(* IEC 61131-3 sources: STEPROBOT/docs/plc_fixed_job_v1_2/现场升级_20261117, 10 files *)

(* ---- GVL_FileBridge.st ---- *)
{attribute 'qualified_only'}
VAR_GLOBAL PERSISTENT RETAIN
    (* Reserve these MW ranges in the FIELD project before importing. *)
    aCommand AT %MW6000 : ARRAY[0..119] OF WORD;
    aHeartbeat AT %MW6120 : ARRAY[0..4] OF WORD;
    aStatus AT %MW6200 : ARRAY[0..63] OF WORD;
END_VAR
VAR_GLOBAL
    (* LOCAL configuration only. Never map credentials/permit to Modbus. *)
    xFileTransferPermit : BOOL := FALSE;
    xReset : BOOL := FALSE;
    sFtpUser : STRING(64) := '';
    sFtpPassword : STRING(64) := '';
    aBuffer : ARRAY[0..1048575] OF BYTE;
    (* One-time LOCAL commissioning: exact existing project already bound to these three GDI numbers.
       This mode reuses bindings. It never edits robot system configuration. *)
    xFixedMappingConfirmed : BOOL := TRUE;
    sFixedProject : STRING(64) := 'pcjob_20261116_201104_7f547f98.sr';
    uiFixedCapture : UINT := UINT#1;
    uiFixedPath : UINT := UINT#2;
    uiFixedReturn : UINT := UINT#3;
    (* Nonretained: a reboot or failed update never authorizes a partly updated project. *)
    xFixedUpdateBusy : BOOL;
    xFixedReady : BOOL;
    xFixedIdle : BOOL;
END_VAR

(* ---- GVL_FileBridgeRetain.st ---- *)
{attribute 'qualified_only'}
VAR_GLOBAL PERSISTENT RETAIN
    udiBootCounter : UDINT := UDINT#0;
END_VAR

(* ---- GVL_RobotBridge.st ---- *)
{attribute 'qualified_only'}
VAR_GLOBAL PERSISTENT RETAIN
    // PC <-> PLC. Inovance native Modbus TCP slave: MWn <-> HR offset n.
    // Commission by reading HR300=16#4D42 and HR301=2 before permitting motion.
    aHostCmd AT %MW200 : ARRAY[0..15] OF WORD;
    aHostStatus AT %MW300 : ARRAY[0..63] OF WORD;

END_VAR

VAR_GLOBAL
    // PLC master -> STEP slave: FC04 / offset 0 / 32 WORD.
    aRobotRx : ARRAY[0..31] OF WORD;
    // PLC master -> STEP slave: ONE FC16 / offset 0 / 2 WORDs.
    // Map BOTH aRobotTx[0] and aRobotTx[1], NOT wRobotTxControl alone.
    aRobotTx : ARRAY[0..1] OF WORD;
    wRobotTxControl : WORD; // first-word diagnostic alias, not a separate channel

    // Local commissioning/operation inputs. Do not map these into aHostCmd.
    xCommissioned : BOOL := FALSE;
    // Set locally ONLY after checking DI49..56 and the GDI program bindings.
    xGdiProgramMappingConfirmed : BOOL := FALSE;
    xRemotePermit : BOOL := FALSE;
    // Optional native master/channel fault. FALSE leaves DO42 watchdog in use.
    xNativeModbusError : BOOL := FALSE;

    // Published live diagnostics.
    xRobotLinkOK : BOOL;
    xRobotRunning : BOOL;
    xRobotPaused : BOOL;
    xRobotStopped : BOOL;
    xRobotEnabled : BOOL;
    xRobotAlarm : BOOL;
    xRobotEmergency : BOOL;
    xRobotExternalAuto : BOOL;
    xHostRegistered : BOOL;
    xHostAlive : BOOL;
    xBusy : BOOL;
    xStopInterlock : BOOL;
    xLoadOperatorConfirmed : BOOL;
    uiFixedJobGuardVersion : UINT;
END_VAR

(* ---- GVL_RobotBridgeRetain.st ---- *)
{attribute 'qualified_only'}
VAR_GLOBAL PERSISTENT RETAIN
    // Incremented on application initialization, not on every scan.
    // Also require a fresh registration; a cold reset can reset RETAIN memory.
    udiBootCounter : UDINT := 0;
END_VAR

(* ---- F_FileCrc32.st ---- *)
FUNCTION F_FileCrc32 : UDINT
VAR_INPUT
    pData : POINTER TO BYTE;
    uiCount : UINT;
    udiSeed : UDINT;
END_VAR
VAR
    udiCrc : UDINT;
    uiI : UINT;
    uiBit : UINT;
END_VAR
(* Running reflected CRC-32. Caller supplies initial FFFFFFFF and final XOR. *)
udiCrc := udiSeed;
IF uiCount > UINT#0 THEN
    FOR uiI := UINT#0 TO uiCount - UINT#1 DO
        udiCrc := udiCrc XOR BYTE_TO_UDINT(pData[uiI]);
        FOR uiBit := UINT#0 TO UINT#7 DO
            IF (udiCrc AND UDINT#1) <> UDINT#0 THEN
                udiCrc := SHR(udiCrc, 1) XOR UDINT#16#EDB88320;
            ELSE
                udiCrc := SHR(udiCrc, 1);
            END_IF;
        END_FOR;
    END_FOR;
END_IF;
F_FileCrc32 := udiCrc;
END_FUNCTION

(* ---- F_FileNameValid.st ---- *)
FUNCTION F_FileNameValid : BOOL
VAR_INPUT
    sName : STRING(64);
    xProject : BOOL;
END_VAR
VAR
    pName : POINTER TO BYTE;
    uiI : UINT;
    uiBaseLength : UINT;
    xValid : BOOL;
    xChar : BOOL;
END_VAR
(* Flat lowercase ASCII names; no slash, CR/LF, spaces, or extra dots. *)
xValid := FALSE;
uiBaseLength := UINT#0;
IF xProject THEN
    IF (LEFT(sName, 6) = 'pcjob_') AND (RIGHT(sName, 3) = '.sr')
        AND (LEN(sName) >= 12) AND (LEN(sName) <= 48) THEN
        uiBaseLength := INT_TO_UINT(LEN(sName)) - UINT#3;
    END_IF;
ELSE
    IF (LEN(sName) >= 5) AND (LEN(sName) <= 48) THEN
        IF (RIGHT(sName, 4) = '.srp') OR (RIGHT(sName, 4) = '.srd')
            OR (RIGHT(sName, 4) = '.txt') THEN
            uiBaseLength := INT_TO_UINT(LEN(sName)) - UINT#4;
        END_IF;
    END_IF;
END_IF;
IF uiBaseLength > UINT#0 THEN
    xValid := TRUE;
    pName := ADR(sName);
    FOR uiI := UINT#0 TO uiBaseLength - UINT#1 DO
        xChar := ((pName[uiI] >= BYTE#97) AND (pName[uiI] <= BYTE#122))
            OR ((pName[uiI] >= BYTE#48) AND (pName[uiI] <= BYTE#57))
            OR (pName[uiI] = BYTE#95);
        IF NOT xChar THEN xValid := FALSE; END_IF;
    END_FOR;
END_IF;
F_FileNameValid := xValid;
END_FUNCTION

(* ---- F_FixedFileValid.st ---- *)
FUNCTION F_FixedFileValid : BOOL
VAR_INPUT
    sName : STRING(64);
END_VAR
F_FixedFileValid := (sName = '_project.srd')
    OR (sName = 'capture_home.srp') OR (sName = 'capture_home.srd')
    OR (sName = 'helix_25mms.srp') OR (sName = 'helix_25mms.srd')
    OR (sName = 'go_home.srp') OR (sName = 'go_home.srd');
END_FUNCTION

(* ---- FB_FileFtp.st ---- *)
FUNCTION_BLOCK FB_FileFtp
VAR_INPUT
    xStart : BOOL;
    xAbort : BOOL;
    pBuffer : POINTER TO BYTE;
    udiSize : UDINT;
    sProject : STRING(64);
    sFile : STRING(64);
    xCreateProject : BOOL;
    xReplaceFixed : BOOL;
    sUser : STRING(64);
    sPassword : STRING(64);
END_VAR
VAR CONSTANT
    cdiControlID : DINT := DINT#245;
    cdiDataID : DINT := DINT#246;
END_VAR
VAR_OUTPUT
    xDone : BOOL := FALSE;
    xTestPassed : BOOL := FALSE;
    xError : BOOL := FALSE;
    xLoginOk : BOOL := FALSE;
    xBaseDirOk : BOOL := FALSE;
    xScratchCreated : BOOL := FALSE;
    xUploadComplete : BOOL := FALSE;
    xReadbackComplete : BOOL := FALSE;
    xContentMatch : BOOL := FALSE;
    xQuitOk : BOOL := FALSE;
    xCleanupOk : BOOL := FALSE;
    uiStep : UINT := UINT#0;
    uiErrorStage : UINT := UINT#0;
    wErrorID : WORD := WORD#0;
    wDataCloseErrorID : WORD := WORD#0;
    wControlCloseErrorID : WORD := WORD#0;
    udiExpectedBytes : UDINT := UDINT#0;
    udiUploadedBytes : UDINT := UDINT#0;
    udiReadbackBytes : UDINT := UDINT#0;
    uiReplyCode : UINT := UINT#0;
    uiUserReplyCode : UINT := UINT#0;
    uiPassReplyCode : UINT := UINT#0;
    uiBaseDirReplyCode : UINT := UINT#0;
    uiNameCheckReplyCode : UINT := UINT#0;
    uiMkdReplyCode : UINT := UINT#0;
    uiStorReplyCode : UINT := UINT#0;
    uiUploadCompleteCode : UINT := UINT#0;
    uiRetrReplyCode : UINT := UINT#0;
    uiDownloadCompleteCode : UINT := UINT#0;
    uiPasvPort : UINT := UINT#0;
    wReadbackEndStatus : WORD := WORD#0;
    sRemotePath : STRING(160);
    sLastReply : STRING(255);
    sMkdReply : STRING(255);
    sPasvReply : STRING(255);
    sUploadReply : STRING(255);
    sDownloadReply : STRING(255);
    xControlOwned : BOOL := FALSE;
    xDataOwned : BOOL := FALSE;
    xUploadDataConnected : BOOL := FALSE;
    xDownloadDataConnected : BOOL := FALSE;
    xLineTruncated : BOOL := FALSE;

END_VAR
VAR
    (* Caller owns immutable buffer until xDone and clean socket closure. *)
    xAbortLatched : BOOL;
    xProgress : BOOL;
    xDirectoryReady : BOOL;
    xReplaceRun : BOOL;
    sFileRun : STRING(64);
    pBufferRun : POINTER TO BYTE;

    stControlServer : CmpHCTCPIP.ADDRESS := (strIPAddr := '192.168.3.188', uiPort := UINT#21);
    stDataServer : CmpHCTCPIP.ADDRESS;
    fbControlClient : CmpHCTCPIP.SktTCPClient;
    fbControlReceive : CmpHCTCPIP.SktTCPRecv;
    fbControlSend : CmpHCTCPIP.SktTCPSend;
    fbControlClose : CmpHCTCPIP.SktClose;
    fbDataClient : CmpHCTCPIP.SktTCPClient;
    fbDataSend : CmpHCTCPIP.SktTCPSend;
    fbDataReceive : CmpHCTCPIP.SktTCPRecv;
    fbDataClose : CmpHCTCPIP.SktClose;
    fbReplyTimeout : TON;
    fbCommandTimeout : TON;
    fbUploadTimeout : TON;
    fbReadbackTimeout : TON;
    fbDataCloseTimeout : TON;
    fbControlCloseTimeout : TON;

    xStartOld : BOOL := FALSE;
    xFail : BOOL := FALSE;
    xFinishedNow : BOOL := FALSE;
    wPendingError : WORD := WORD#0;
    uiPendingStage : UINT := UINT#0;
    uiPhase : UINT := UINT#0;
    uiNextCommand : UINT := UINT#0;
    uiTransferMode : UINT := UINT#0;
    xReplyReady : BOOL := FALSE;
    xReplyAccepted : BOOL := FALSE;
    xDigits : BOOL := FALSE;
    xMultiline : BOOL := FALSE;
    sMultilineCode : STRING(3);
    sLine : STRING(255);
    pLine : POINTER TO BYTE;
    uiLineLength : UINT := UINT#0;
    aControlRx : ARRAY[0..0] OF BYTE;
    sCommand : STRING(160);
    pCommand : POINTER TO BYTE;
    uiCommandIndex : UINT := UINT#0;
    uiCommandLength : UINT := UINT#0;
    aControlTx : ARRAY[0..0] OF BYTE;
    aDataTx : ARRAY[0..0] OF BYTE;
    aDataRx : ARRAY[0..0] OF BYTE;
    sUserRun : STRING(64);
    sPasswordRun : STRING(64);
    sScratchRun : STRING(64);
    pCredential : POINTER TO BYTE;
    uiI : UINT := UINT#0;
    xNameCharacter : BOOL := FALSE;
    xBytesMatch : BOOL := FALSE;
    xReadbackEndCandidate : BOOL := FALSE;
    xDataCloseFailed : BOOL := FALSE;
    pReply : POINTER TO BYTE;
    aPasv : ARRAY[0..5] OF UINT;
    uiPasvField : UINT := UINT#0;
    uiPasvValue : UINT := UINT#0;
    xPasvValid : BOOL := FALSE;
    xPasvInTuple : BOOL := FALSE;
    xPasvClosed : BOOL := FALSE;
    xPasvHasDigit : BOOL := FALSE;
END_VAR
(* Derived from field-passed PRG_FtpUploadProbe. New bridge is NOT field validated. *)
(* IDs 245/246 must be free; default cabinet 192.168.3.188:21. *)
(* One-byte send/reset preserves the tested Socket behavior. No motion commands. *)
pLine := ADR(sLine);
pCommand := ADR(sCommand);
xFail := FALSE;
xFinishedNow := FALSE;
xReplyReady := FALSE;
wPendingError := WORD#0;
uiPendingStage := UINT#20 + uiPhase * UINT#10;

IF uiStep = UINT#40 THEN
    aControlTx[0] := pCommand[uiCommandIndex];
END_IF;
IF uiStep = UINT#60 THEN
    IF udiUploadedBytes < udiExpectedBytes THEN
        aDataTx[0] := pBufferRun[udiUploadedBytes];
    END_IF;
END_IF;

fbControlClient(xExecute := uiStep = UINT#10, diConnectID := cdiControlID,
    stServerAddress := stControlServer);
fbControlReceive(xEnable := uiStep = UINT#20, diConnectID := cdiControlID,
    abyData := aControlRx, uiDataSize := UINT#1);
fbControlSend(xExecute := uiStep = UINT#40, diConnectID := cdiControlID,
    abyData := aControlTx, uiDataSize := UINT#1, uiTimeOut := UINT#1000);
fbDataClient(xExecute := uiStep = UINT#50, diConnectID := cdiDataID,
    stServerAddress := stDataServer);
fbDataSend(xExecute := uiStep = UINT#60, diConnectID := cdiDataID,
    abyData := aDataTx, uiDataSize := UINT#1, uiTimeOut := UINT#1000);
fbDataReceive(xEnable := uiStep = UINT#70, diConnectID := cdiDataID,
    abyData := aDataRx, uiDataSize := UINT#1);
fbDataClose(xExecute := ((uiStep = UINT#80) OR (uiStep = UINT#90))
    AND xDataOwned AND NOT xDataCloseFailed, diConnectID := cdiDataID);
fbControlClose(xExecute := (uiStep = UINT#95) AND xControlOwned,
    diConnectID := cdiControlID);
fbReplyTimeout(IN := uiStep = UINT#20, PT := T#20s);
fbCommandTimeout(IN := (uiStep = UINT#40) OR (uiStep = UINT#45), PT := T#30s);
xProgress := ((uiStep = UINT#60) AND fbDataSend.xDone)
    OR ((uiStep = UINT#70) AND (fbDataReceive.uiCount > UINT#0));
fbUploadTimeout(IN := ((uiStep = UINT#60) OR (uiStep = UINT#65)) AND NOT xProgress,
    PT := T#30s);
fbReadbackTimeout(IN := (uiStep = UINT#70) AND NOT xProgress, PT := T#30s);
fbDataCloseTimeout(IN := ((uiStep = UINT#80) OR (uiStep = UINT#90))
    AND xDataOwned AND NOT xDataCloseFailed, PT := T#5s);
fbControlCloseTimeout(IN := uiStep = UINT#95, PT := T#5s);

(* Bounded control-reply parser; identical-code SPACE terminates multiline replies. *)
IF (uiStep = UINT#20) AND NOT fbControlReceive.xError THEN
    IF fbControlReceive.uiCount > UINT#0 THEN
        IF aControlRx[0] = BYTE#10 THEN
            IF uiLineLength > UINT#0 THEN
                IF pLine[uiLineLength - UINT#1] = BYTE#13 THEN
                    uiLineLength := uiLineLength - UINT#1;
                    pLine[uiLineLength] := BYTE#0;
                END_IF;
            END_IF;
            IF xMultiline THEN
                IF LEFT(sLine, 4) = CONCAT(sMultilineCode, ' ') THEN
                    xMultiline := FALSE;
                    xReplyReady := TRUE;
                END_IF;
            ELSE
                xDigits := FALSE;
                IF uiLineLength >= UINT#4 THEN
                    xDigits := (pLine[0] >= BYTE#48) AND (pLine[0] <= BYTE#57)
                        AND (pLine[1] >= BYTE#48) AND (pLine[1] <= BYTE#57)
                        AND (pLine[2] >= BYTE#48) AND (pLine[2] <= BYTE#57);
                END_IF;
                IF xDigits THEN
                    IF pLine[3] = BYTE#45 THEN
                        xMultiline := TRUE;
                        sMultilineCode := LEFT(sLine, 3);
                    ELSIF pLine[3] = BYTE#32 THEN
                        xReplyReady := TRUE;
                    ELSE
                        xFail := TRUE;
                        wPendingError := WORD#16#F203;
                    END_IF;
                ELSE
                    xFail := TRUE;
                    wPendingError := WORD#16#F203;
                END_IF;
            END_IF;
            IF xReplyReady THEN
                uiReplyCode := (BYTE_TO_UINT(pLine[0]) - UINT#48) * UINT#100
                    + (BYTE_TO_UINT(pLine[1]) - UINT#48) * UINT#10
                    + BYTE_TO_UINT(pLine[2]) - UINT#48;
                sLastReply := sLine;
            ELSIF xFail THEN
                sLastReply := sLine;
            END_IF;
            sLine := '';
            uiLineLength := UINT#0;
        ELSE
            IF uiLineLength < UINT#255 THEN
                pLine[uiLineLength] := aControlRx[0];
                uiLineLength := uiLineLength + UINT#1;
                pLine[uiLineLength] := BYTE#0;
            ELSE
                xLineTruncated := TRUE;
                sLastReply := sLine;
                xFail := TRUE;
                wPendingError := WORD#16#F204;
            END_IF;
        END_IF;
    END_IF;
END_IF;

CASE uiStep OF
    UINT#0:
        IF xStart AND NOT xStartOld THEN
            xAbortLatched := FALSE;
            xDirectoryReady := FALSE;
            xDone := FALSE;
            xTestPassed := FALSE;
            xError := FALSE;
            xLoginOk := FALSE;
            xBaseDirOk := FALSE;
            xScratchCreated := FALSE;
            xUploadComplete := FALSE;
            xReadbackComplete := FALSE;
            xContentMatch := FALSE;
            xQuitOk := FALSE;
            xCleanupOk := FALSE;
            xUploadDataConnected := FALSE;
            xDownloadDataConnected := FALSE;
            xDataCloseFailed := FALSE;
            xLineTruncated := FALSE;
            xReadbackEndCandidate := FALSE;
            xBytesMatch := TRUE;
            uiErrorStage := UINT#0;
            wErrorID := WORD#0;
            wDataCloseErrorID := WORD#0;
            wControlCloseErrorID := WORD#0;
            wReadbackEndStatus := WORD#0;
            udiUploadedBytes := UDINT#0;
            udiReadbackBytes := UDINT#0;
            uiReplyCode := UINT#0;
            uiUserReplyCode := UINT#0;
            uiPassReplyCode := UINT#0;
            uiBaseDirReplyCode := UINT#0;
            uiNameCheckReplyCode := UINT#0;
            uiMkdReplyCode := UINT#0;
            uiStorReplyCode := UINT#0;
            uiUploadCompleteCode := UINT#0;
            uiRetrReplyCode := UINT#0;
            uiDownloadCompleteCode := UINT#0;
            uiPasvPort := UINT#0;
            sLastReply := '';
            sMkdReply := '';
            sPasvReply := '';
            sUploadReply := '';
            sDownloadReply := '';
            sLine := '';
            uiLineLength := UINT#0;
            xMultiline := FALSE;
            sMultilineCode := '';
            uiPhase := UINT#0;
            uiTransferMode := UINT#0;
            sUserRun := sUser;
            sPasswordRun := sPassword;
            sScratchRun := sProject;
            sFileRun := sFile;
            xReplaceRun := xReplaceFixed;
            pBufferRun := pBuffer;
            sRemotePath := CONCAT(CONCAT(CONCAT('/UserPrograms/', sScratchRun), '/'), sFileRun);
            udiExpectedBytes := udiSize;
            uiPendingStage := UINT#1;
            IF (LEN(sUserRun) = 0) OR (LEN(sPasswordRun) = 0) THEN
                xFail := TRUE;
                wPendingError := WORD#16#F200;
            ELSE
                pCredential := ADR(sUserRun);
                FOR uiI := UINT#0 TO INT_TO_UINT(LEN(sUserRun)) - UINT#1 DO
                    IF (pCredential[uiI] < BYTE#32) OR (pCredential[uiI] > BYTE#126) THEN
                        xFail := TRUE;
                        wPendingError := WORD#16#F207;
                    END_IF;
                END_FOR;
                pCredential := ADR(sPasswordRun);
                FOR uiI := UINT#0 TO INT_TO_UINT(LEN(sPasswordRun)) - UINT#1 DO
                    IF (pCredential[uiI] < BYTE#32) OR (pCredential[uiI] > BYTE#126) THEN
                        xFail := TRUE;
                        wPendingError := WORD#16#F207;
                    END_IF;
                END_FOR;
            END_IF;
            IF NOT F_FileNameValid(sScratchRun, TRUE)
                OR NOT F_FileNameValid(sFileRun, FALSE)
                OR (udiExpectedBytes > UDINT#1048576)
                OR (pBufferRun = 0) THEN
                xFail := TRUE;
                wPendingError := WORD#16#F209;
            END_IF;
            IF xReplaceRun AND (NOT GVL_FileBridge.xFixedMappingConfirmed
                OR (GVL_RobotBridge.uiFixedJobGuardVersion <> UINT#120)
                OR NOT GVL_FileBridge.xFixedIdle OR (sScratchRun <> GVL_FileBridge.sFixedProject)
                OR NOT F_FixedFileValid(sFileRun)) THEN
                xFail := TRUE;
                wPendingError := WORD#16#F20C;
            END_IF;
            IF NOT xFail THEN
                uiStep := UINT#10;
            END_IF;
        END_IF;

    UINT#10:
        IF fbControlClient.xError THEN
            xFail := TRUE;
            wPendingError := fbControlClient.wErrorID;
            uiPendingStage := UINT#10;
        ELSIF fbControlClient.xDone THEN
            xControlOwned := TRUE;
            uiStep := UINT#20;
        END_IF;

    UINT#20:
        IF fbControlReceive.xError THEN
            xFail := TRUE;
            wPendingError := fbControlReceive.wErrorID;
        ELSIF NOT xFail THEN
            IF xReplyReady THEN
                xReplyAccepted := FALSE;
                CASE uiPhase OF
                    UINT#0:
                        IF uiReplyCode = UINT#220 THEN
                            xReplyAccepted := TRUE;
                            uiNextCommand := UINT#1;
                            uiStep := UINT#30;
                        ELSIF uiReplyCode = UINT#120 THEN
                            xReplyAccepted := TRUE;
                        END_IF;
                    UINT#1:
                        uiUserReplyCode := uiReplyCode;
                        IF uiReplyCode = UINT#331 THEN
                            xReplyAccepted := TRUE;
                            uiNextCommand := UINT#2;
                            uiStep := UINT#30;
                        ELSIF uiReplyCode = UINT#230 THEN
                            xReplyAccepted := TRUE;
                            xLoginOk := TRUE;
                            uiNextCommand := UINT#3;
                            uiStep := UINT#30;
                        END_IF;
                    UINT#2:
                        uiPassReplyCode := uiReplyCode;
                        IF uiReplyCode = UINT#230 THEN
                            xReplyAccepted := TRUE;
                            xLoginOk := TRUE;
                            uiNextCommand := UINT#3;
                            uiStep := UINT#30;
                        END_IF;
                    UINT#3:
                        uiBaseDirReplyCode := uiReplyCode;
                        IF uiReplyCode = UINT#250 THEN
                            xReplyAccepted := TRUE;
                            xBaseDirOk := TRUE;
                            IF xCreateProject OR xReplaceRun THEN
                                uiNextCommand := UINT#14;
                            ELSE
                                uiNextCommand := UINT#5;
                            END_IF;
                            uiStep := UINT#30;
                        END_IF;
                    UINT#14:
                        uiNameCheckReplyCode := uiReplyCode;
                        IF uiReplyCode = UINT#550 THEN
                            xReplyAccepted := TRUE;
                            IF xReplaceRun THEN
                                (* Fixed binding must already exist: never silently create another target. *)
                                xFail := TRUE;
                                wPendingError := WORD#16#F20B;
                            ELSE
                                uiNextCommand := UINT#4;
                                uiStep := UINT#30;
                            END_IF;
                        ELSIF uiReplyCode = UINT#250 THEN
                            xReplyAccepted := TRUE;
                            IF xReplaceRun THEN
                                xDirectoryReady := TRUE;
                                uiNextCommand := UINT#6;
                                uiStep := UINT#30;
                            ELSE
                                (* Original mode retains its no-overwrite behavior. *)
                                xFail := TRUE;
                                wPendingError := WORD#16#F208;
                            END_IF;
                        END_IF;
                    UINT#4:
                        uiMkdReplyCode := uiReplyCode;
                        sMkdReply := sLastReply;
                        IF uiReplyCode = UINT#257 THEN
                            xReplyAccepted := TRUE;
                            xScratchCreated := TRUE;
                            uiNextCommand := UINT#5;
                            uiStep := UINT#30;
                        END_IF;
                    UINT#5:
                        IF uiReplyCode = UINT#250 THEN
                            xDirectoryReady := TRUE;
                            xReplyAccepted := TRUE;
                            uiNextCommand := UINT#6;
                            uiStep := UINT#30;
                        END_IF;
                    UINT#6:
                        IF uiReplyCode = UINT#200 THEN
                            xReplyAccepted := TRUE;
                            uiNextCommand := UINT#7;
                            uiStep := UINT#30;
                        END_IF;
                    UINT#7, UINT#10:
                        IF uiReplyCode = UINT#227 THEN
                            xReplyAccepted := TRUE;
                            sPasvReply := sLastReply;
                            uiStep := UINT#35;
                        END_IF;
                    UINT#8:
                        uiStorReplyCode := uiReplyCode;
                        IF (uiReplyCode = UINT#125) OR (uiReplyCode = UINT#150) THEN
                            xReplyAccepted := TRUE;
                            IF udiExpectedBytes = UDINT#0 THEN
                                (* Empty STOR still needs data EOF, 226 and exact RETR. *)
                                uiStep := UINT#80;
                            ELSE
                                uiStep := UINT#60;
                            END_IF;
                        END_IF;
                    UINT#9:
                        uiUploadCompleteCode := uiReplyCode;
                        sUploadReply := sLastReply;
                        IF (uiReplyCode = UINT#226) OR (uiReplyCode = UINT#250) THEN
                            xReplyAccepted := TRUE;
                            xUploadComplete := TRUE;
                            uiNextCommand := UINT#10;
                            uiStep := UINT#30;
                        END_IF;
                    UINT#11:
                        uiRetrReplyCode := uiReplyCode;
                        IF (uiReplyCode = UINT#125) OR (uiReplyCode = UINT#150) THEN
                            xReplyAccepted := TRUE;
                            uiStep := UINT#70;
                        END_IF;
                    UINT#12:
                        uiDownloadCompleteCode := uiReplyCode;
                        sDownloadReply := sLastReply;
                        IF (uiReplyCode = UINT#226) OR (uiReplyCode = UINT#250) THEN
                            xReplyAccepted := TRUE;
                            xReadbackComplete := TRUE;
                            xContentMatch := xBytesMatch AND xReadbackEndCandidate
                                AND (udiReadbackBytes = udiExpectedBytes);
                            IF xContentMatch THEN
                                uiNextCommand := UINT#13;
                                uiStep := UINT#30;
                            ELSE
                                xFail := TRUE;
                                wPendingError := WORD#16#F205;
                            END_IF;
                        END_IF;
                    UINT#13:
                        IF uiReplyCode = UINT#221 THEN
                            xReplyAccepted := TRUE;
                            xQuitOk := TRUE;
                            uiStep := UINT#90;
                        END_IF;
                END_CASE;
                IF NOT xReplyAccepted THEN
                    xFail := TRUE;
                    wPendingError := WORD#16#F202;
                END_IF;
            ELSIF fbReplyTimeout.Q THEN
                xFail := TRUE;
                wPendingError := WORD#16#F201;
            END_IF;
        END_IF;

    UINT#30:
        uiPhase := uiNextCommand;
        CASE uiNextCommand OF
            UINT#1: sCommand := CONCAT(CONCAT('USER ', sUserRun), '$R$N');
            UINT#2: sCommand := CONCAT(CONCAT('PASS ', sPasswordRun), '$R$N');
            UINT#3: sCommand := 'CWD /UserPrograms$R$N';
            UINT#4: sCommand := CONCAT(CONCAT('MKD ', sScratchRun), '$R$N');
            UINT#5, UINT#14: sCommand := CONCAT(CONCAT('CWD ', sScratchRun), '$R$N');
            UINT#6: sCommand := 'TYPE I$R$N';
            UINT#7, UINT#10: sCommand := 'PASV$R$N';
            UINT#8: sCommand := CONCAT(CONCAT('STOR ', sFileRun), '$R$N');
            UINT#11: sCommand := CONCAT(CONCAT('RETR ', sFileRun), '$R$N');
            UINT#13: sCommand := 'QUIT$R$N';
        ELSE
            xFail := TRUE;
            wPendingError := WORD#16#F20A;
        END_CASE;
        IF NOT xFail THEN
            uiCommandLength := INT_TO_UINT(LEN(sCommand));
            uiCommandIndex := UINT#0;
            uiStep := UINT#40;
        END_IF;

    UINT#35:
        (* Parse six decimal octets in the first parenthesized PASV tuple. *)
        pReply := ADR(sPasvReply);
        xPasvValid := TRUE;
        xPasvInTuple := FALSE;
        xPasvClosed := FALSE;
        xPasvHasDigit := FALSE;
        uiPasvField := UINT#0;
        uiPasvValue := UINT#0;
        FOR uiI := UINT#0 TO INT_TO_UINT(LEN(sPasvReply)) - UINT#1 DO
            IF NOT xPasvInTuple THEN
                IF pReply[uiI] = BYTE#40 THEN
                    xPasvInTuple := TRUE;
                END_IF;
            ELSIF NOT xPasvClosed THEN
                IF (pReply[uiI] >= BYTE#48) AND (pReply[uiI] <= BYTE#57) THEN
                    xPasvHasDigit := TRUE;
                    IF uiPasvValue <= UINT#255 THEN
                        uiPasvValue := uiPasvValue * UINT#10 + BYTE_TO_UINT(pReply[uiI]) - UINT#48;
                        IF uiPasvValue > UINT#255 THEN
                            xPasvValid := FALSE;
                        END_IF;
                    ELSE
                        xPasvValid := FALSE;
                    END_IF;
                ELSIF (pReply[uiI] = BYTE#44) OR (pReply[uiI] = BYTE#41) THEN
                    IF NOT xPasvHasDigit OR (uiPasvField > UINT#5) OR (uiPasvValue > UINT#255) THEN
                        xPasvValid := FALSE;
                    ELSE
                        aPasv[uiPasvField] := uiPasvValue;
                        uiPasvField := uiPasvField + UINT#1;
                    END_IF;
                    uiPasvValue := UINT#0;
                    xPasvHasDigit := FALSE;
                    IF pReply[uiI] = BYTE#41 THEN
                        xPasvClosed := TRUE;
                    END_IF;
                ELSE
                    xPasvValid := FALSE;
                END_IF;
            END_IF;
        END_FOR;
        IF NOT xPasvInTuple OR NOT xPasvClosed OR (uiPasvField <> UINT#6) THEN
            xPasvValid := FALSE;
        END_IF;
        IF xPasvValid THEN
            uiPasvPort := aPasv[4] * UINT#256 + aPasv[5];
            IF (uiPasvPort = UINT#0) OR (uiPasvPort = UINT#21) THEN
                xPasvValid := FALSE;
            END_IF;
        END_IF;
        IF xPasvValid THEN
            (* Data connections are pinned to the control server, not a third-party PASV IP. *)
            stDataServer.strIPAddr := stControlServer.strIPAddr;
            stDataServer.uiPort := uiPasvPort;
            xDataCloseFailed := FALSE;
            IF uiPhase = UINT#7 THEN
                uiTransferMode := UINT#1;
            ELSE
                uiTransferMode := UINT#2;
            END_IF;
            uiStep := UINT#50;
        ELSE
            xFail := TRUE;
            wPendingError := WORD#16#F20B;
        END_IF;

    UINT#40:
        IF fbControlSend.xError THEN
            xFail := TRUE;
            wPendingError := fbControlSend.wErrorID;
        ELSIF fbControlSend.xDone THEN
            uiCommandIndex := uiCommandIndex + UINT#1;
            uiStep := UINT#45;
        ELSIF fbCommandTimeout.Q THEN
            xFail := TRUE;
            wPendingError := WORD#16#F206;
        END_IF;

    UINT#45:
        IF uiCommandIndex >= uiCommandLength THEN
            sCommand := '';
            aControlTx[0] := BYTE#0;
            sLine := '';
            uiLineLength := UINT#0;
            xMultiline := FALSE;
            sMultilineCode := '';
            uiStep := UINT#20;
        ELSIF fbCommandTimeout.Q THEN
            xFail := TRUE;
            wPendingError := WORD#16#F206;
        ELSE
            uiStep := UINT#40;
        END_IF;

    UINT#50:
        uiPendingStage := UINT#200 + uiTransferMode;
        IF fbDataClient.xError THEN
            xFail := TRUE;
            wPendingError := fbDataClient.wErrorID;
        ELSIF fbDataClient.xDone THEN
            xDataOwned := TRUE;
            IF uiTransferMode = UINT#1 THEN
                xUploadDataConnected := TRUE;
                uiNextCommand := UINT#8;
            ELSE
                xDownloadDataConnected := TRUE;
                uiNextCommand := UINT#11;
            END_IF;
            uiStep := UINT#30;
        END_IF;

    UINT#60:
        uiPendingStage := UINT#210;
        IF fbDataSend.xError THEN
            xFail := TRUE;
            wPendingError := fbDataSend.wErrorID;
        ELSIF fbDataSend.xDone THEN
            udiUploadedBytes := udiUploadedBytes + UDINT#1;
            uiStep := UINT#65;
        ELSIF fbUploadTimeout.Q THEN
            xFail := TRUE;
            wPendingError := WORD#16#F206;
        END_IF;

    UINT#65:
        uiPendingStage := UINT#210;
        IF udiUploadedBytes >= udiExpectedBytes THEN
            aDataTx[0] := BYTE#0;
            uiStep := UINT#80;
        ELSIF fbUploadTimeout.Q THEN
            xFail := TRUE;
            wPendingError := WORD#16#F206;
        ELSE
            uiStep := UINT#60;
        END_IF;

    UINT#70:
        uiPendingStage := UINT#220;
        IF fbDataReceive.xError THEN
            wReadbackEndStatus := fbDataReceive.wErrorID;
            (* In the supplied source, zero-length recv and recv failure share 0011. *)
            (* This is only an end candidate: exact bytes AND FTP completion are required. *)
            IF (wReadbackEndStatus = WORD#16#0011) AND xBytesMatch
                AND (udiReadbackBytes = udiExpectedBytes) THEN
                xReadbackEndCandidate := TRUE;
                uiStep := UINT#80;
            ELSE
                xFail := TRUE;
                wPendingError := fbDataReceive.wErrorID;
            END_IF;
        ELSIF fbDataReceive.uiCount > UINT#0 THEN
            IF udiReadbackBytes >= udiExpectedBytes THEN
                xBytesMatch := FALSE;
                xFail := TRUE;
                wPendingError := WORD#16#F205;
            ELSE
                IF aDataRx[0] <> pBufferRun[udiReadbackBytes] THEN
                    xBytesMatch := FALSE;
                    xFail := TRUE;
                    wPendingError := WORD#16#F205;
                END_IF;
                udiReadbackBytes := udiReadbackBytes + UDINT#1;
            END_IF;
        ELSIF fbReadbackTimeout.Q THEN
            xFail := TRUE;
            wPendingError := WORD#16#F201;
        END_IF;

    UINT#80:
        IF fbDataClose.xError OR fbDataCloseTimeout.Q THEN
            IF fbDataClose.xError THEN
                wDataCloseErrorID := fbDataClose.wErrorID;
            ELSE
                wDataCloseErrorID := WORD#16#F20C;
            END_IF;
            xDataCloseFailed := TRUE;
            IF NOT xError THEN
                xError := TRUE;
                wErrorID := wDataCloseErrorID;
                uiErrorStage := UINT#290;
            END_IF;
            uiStep := UINT#95;
        ELSIF fbDataClose.xDone THEN
            xDataOwned := FALSE;
            IF uiTransferMode = UINT#1 THEN
                uiPhase := UINT#9;
            ELSE
                uiPhase := UINT#12;
            END_IF;
            uiStep := UINT#20;
        END_IF;

    UINT#90:
        IF NOT xDataOwned OR xDataCloseFailed THEN
            uiStep := UINT#95;
        ELSIF fbDataClose.xError OR fbDataCloseTimeout.Q THEN
            IF fbDataClose.xError THEN
                wDataCloseErrorID := fbDataClose.wErrorID;
            ELSE
                wDataCloseErrorID := WORD#16#F20C;
            END_IF;
            xDataCloseFailed := TRUE;
            IF NOT xError THEN
                xError := TRUE;
                wErrorID := wDataCloseErrorID;
                uiErrorStage := UINT#290;
            END_IF;
            uiStep := UINT#95;
        ELSIF fbDataClose.xDone THEN
            xDataOwned := FALSE;
            uiStep := UINT#95;
        END_IF;

    UINT#95:
        IF NOT xControlOwned THEN
            xDone := TRUE;
            xFinishedNow := TRUE;
            uiStep := UINT#100;
        ELSIF fbControlClose.xError OR fbControlCloseTimeout.Q THEN
            IF fbControlClose.xError THEN
                wControlCloseErrorID := fbControlClose.wErrorID;
            ELSE
                wControlCloseErrorID := WORD#16#F20C;
            END_IF;
            IF NOT xError THEN
                xError := TRUE;
                wErrorID := wControlCloseErrorID;
                uiErrorStage := UINT#295;
            END_IF;
            xDone := TRUE;
            xFinishedNow := TRUE;
            uiStep := UINT#100;
        ELSIF fbControlClose.xDone THEN
            xControlOwned := FALSE;
            xDone := TRUE;
            xFinishedNow := TRUE;
            uiStep := UINT#100;
        END_IF;

    UINT#100:
        IF NOT xStart AND NOT xControlOwned AND NOT xDataOwned THEN
            uiStep := UINT#0;
        END_IF;
END_CASE;

(* Never cancel a pending native connect before its terminal result. *)
IF xAbort AND (uiStep <> UINT#0) AND (uiStep <> UINT#100) THEN
    xAbortLatched := TRUE;
END_IF;
IF xAbortLatched AND (uiStep <> UINT#0) AND (uiStep <> UINT#10)
    AND (uiStep <> UINT#50) AND (uiStep <> UINT#90)
    AND (uiStep <> UINT#95) AND (uiStep <> UINT#100) THEN
    xFail := TRUE;
    wPendingError := WORD#16#F20D;
END_IF;
IF xFail THEN
    IF NOT xError THEN
        xError := TRUE;
        wErrorID := wPendingError;
        uiErrorStage := uiPendingStage;
    END_IF;
    uiStep := UINT#90;
END_IF;

IF xFinishedNow THEN
    xCleanupOk := NOT xControlOwned AND NOT xDataOwned
        AND (wDataCloseErrorID = WORD#0) AND (wControlCloseErrorID = WORD#0);
    xTestPassed := xLoginOk AND xBaseDirOk AND xDirectoryReady
        AND xUploadDataConnected AND xDownloadDataConnected
        AND xUploadComplete AND xReadbackComplete AND xContentMatch
        AND xQuitOk AND xCleanupOk AND NOT xError;
    sPasswordRun := '';
    sUserRun := '';
    sCommand := '';
    aControlTx[0] := BYTE#0;
    aDataTx[0] := BYTE#0;
END_IF;
xStartOld := xStart;
END_FUNCTION_BLOCK

(* ---- PRG_FileBridge.st ---- *)
PROGRAM PRG_FileBridge
VAR
    xInit : BOOL;
    xResetOld : BOOL;
    aPrevious : ARRAY[0..119] OF WORD;
    aSeen : ARRAY[0..119] OF WORD;
    aFrame : ARRAY[0..119] OF WORD;
    aAccepted : ARRAY[0..119] OF WORD;
    aFrameBytes : ARRAY[0..235] OF BYTE;
    aPayload : ARRAY[0..191] OF BYTE;
    aNames : ARRAY[0..31] OF STRING(64);
    uiState : UINT;
    wError : WORD;
    udiOwner : UDINT;
    udiAck : UDINT;
    uiAckOp : UINT;
    udiSize : UDINT;
    udiReceived : UDINT;
    udiExpectedCrc : UDINT;
    udiRunningCrc : UDINT := UDINT#16#FFFFFFFF;
    udiTotalSize : UDINT;
    uiVerified : UINT;
    uiExpectedFiles : UINT;
    uiOrdinal : UINT;
    uiMode : UINT;
    sProject : STRING(64);
    sFile : STRING(64);
    fbFtp : FB_FileFtp;
    fbLease : TON;
    wHeartbeatOld : WORD;
    xKick : BOOL;
    xStable : BOOL;
    xNew : BOOL;
    xSame : BOOL;
    xAccept : BOOL;
    xActive : BOOL;
    xClean : BOOL;
    xFileVerified : BOOL;
    xFtpStarted : BOOL;
    wReject : WORD;
    udiRejectSeq : UDINT;
    udiRejectOwner : UDINT;
    wRequestError : WORD;
    udiSeq : UDINT;
    udiSession : UDINT;
    udiBoot : UDINT;
    udiFrameCrc : UDINT;
    udiFrameSize : UDINT;
    udiOffset : UDINT;
    udiFileCrc : UDINT;
    uiOp : UINT;
    uiLength : UINT;
    uiCount : UINT;
    uiIndex : UINT;
    uiField : UINT;
    uiPos : UINT;
    uiI : UINT;
    uiJ : UINT;
    uiSnapshot : UINT;
    wFlags : WORD;
    sNewProject : STRING(64);
    sNewFile : STRING(64);
    pName : POINTER TO BYTE;
    xNamesOk : BOOL;
    xPairsOk : BOOL;
    xFound : BOOL;
    xGlobal : BOOL;
    uiPrograms : UINT;
    sPair : STRING(64);
    sReadyProject : STRING(64);
    uiReadyCapture : UINT;
    uiReadyPath : UINT;
    uiReadyReturn : UINT;
    xFixedConfig : BOOL;
    udiFixedProjectCrc : UDINT;
    uiSessionCapture : UINT;
    uiSessionPath : UINT;
    uiSessionReturn : UINT;
END_VAR

(* This program NEVER writes robot motion/control outputs or GDI selection. *)
IF NOT xInit THEN
    GVL_FileBridge.xFixedReady := FALSE;
    GVL_FileBridge.xFixedUpdateBusy := FALSE;
    IF GVL_FileBridgeRetain.udiBootCounter = UDINT#16#FFFFFFFF THEN
        GVL_FileBridgeRetain.udiBootCounter := UDINT#1;
    ELSE
        GVL_FileBridgeRetain.udiBootCounter := GVL_FileBridgeRetain.udiBootCounter + UDINT#1;
    END_IF;
    FOR uiI := UINT#0 TO UINT#119 DO
        aPrevious[uiI] := GVL_FileBridge.aCommand[uiI];
        aSeen[uiI] := GVL_FileBridge.aCommand[uiI];
    END_FOR;
    xInit := TRUE;
END_IF;

xFixedConfig := GVL_FileBridge.xFixedMappingConfirmed
    AND (GVL_RobotBridge.uiFixedJobGuardVersion = UINT#120)
    AND F_FileNameValid(GVL_FileBridge.sFixedProject, TRUE)
    AND (GVL_FileBridge.uiFixedCapture >= UINT#1) AND (GVL_FileBridge.uiFixedCapture <= UINT#255)
    AND (GVL_FileBridge.uiFixedPath >= UINT#1) AND (GVL_FileBridge.uiFixedPath <= UINT#255)
    AND (GVL_FileBridge.uiFixedReturn >= UINT#1) AND (GVL_FileBridge.uiFixedReturn <= UINT#255)
    AND (GVL_FileBridge.uiFixedCapture <> GVL_FileBridge.uiFixedPath)
    AND (GVL_FileBridge.uiFixedCapture <> GVL_FileBridge.uiFixedReturn)
    AND (GVL_FileBridge.uiFixedPath <> GVL_FileBridge.uiFixedReturn);
GVL_FileBridge.xFixedIdle := GVL_RobotBridge.xRobotLinkOK AND GVL_RobotBridge.xRobotStopped
    AND NOT GVL_RobotBridge.xRobotRunning AND NOT GVL_RobotBridge.xRobotPaused
    AND NOT GVL_RobotBridge.xRobotEnabled AND NOT GVL_RobotBridge.xBusy;
IF NOT xFixedConfig OR (sReadyProject <> GVL_FileBridge.sFixedProject)
    OR (uiReadyCapture <> GVL_FileBridge.uiFixedCapture) OR (uiReadyPath <> GVL_FileBridge.uiFixedPath)
    OR (uiReadyReturn <> GVL_FileBridge.uiFixedReturn) THEN
    GVL_FileBridge.xFixedReady := FALSE;
END_IF;
udiFixedProjectCrc := F_FileCrc32(ADR(GVL_FileBridge.sFixedProject),
    INT_TO_UINT(LEN(GVL_FileBridge.sFixedProject)), UDINT#16#FFFFFFFF) XOR UDINT#16#FFFFFFFF;

xClean := NOT fbFtp.xControlOwned AND NOT fbFtp.xDataOwned
    AND ((fbFtp.uiStep = UINT#0) OR (fbFtp.uiStep = UINT#100));
IF GVL_FileBridge.xReset AND NOT xResetOld AND xClean
    AND (uiState <> UINT#300) AND (uiState <> UINT#310) THEN
    uiState := UINT#0;
    wError := WORD#0;
    udiOwner := UDINT#0;
    udiAck := UDINT#0;
    uiAckOp := UINT#0;
    uiVerified := UINT#0;
    uiExpectedFiles := UINT#0;
    udiReceived := UDINT#0;
    udiSize := UDINT#0;
    xFileVerified := FALSE;
    GVL_FileBridge.xFixedReady := FALSE;
    wReject := WORD#0;
END_IF;
xResetOld := GVL_FileBridge.xReset;

xActive := (uiState = UINT#100) OR (uiState = UINT#200)
    OR (uiState = UINT#300) OR (uiState = UINT#310);
xKick := FALSE;
IF (GVL_FileBridge.aHeartbeat[0] = UDINT_TO_WORD(SHR(udiOwner, 16)))
    AND (GVL_FileBridge.aHeartbeat[1] = UDINT_TO_WORD(udiOwner))
    AND (GVL_FileBridge.aHeartbeat[2] = UDINT_TO_WORD(SHR(GVL_FileBridgeRetain.udiBootCounter, 16)))
    AND (GVL_FileBridge.aHeartbeat[3] = UDINT_TO_WORD(GVL_FileBridgeRetain.udiBootCounter))
    AND (GVL_FileBridge.aHeartbeat[4] <> wHeartbeatOld) THEN
    wHeartbeatOld := GVL_FileBridge.aHeartbeat[4];
    xKick := TRUE;
END_IF;
fbLease(IN := xActive AND NOT xKick, PT := T#10s);

(* Two consecutive identical samples, then CRC of big-endian WORD bytes. *)
xStable := TRUE;
xNew := FALSE;
FOR uiI := UINT#0 TO UINT#119 DO
    aFrame[uiI] := GVL_FileBridge.aCommand[uiI];
    IF aFrame[uiI] <> aPrevious[uiI] THEN xStable := FALSE; END_IF;
    IF aFrame[uiI] <> aSeen[uiI] THEN xNew := TRUE; END_IF;
    aPrevious[uiI] := aFrame[uiI];
END_FOR;
IF xStable AND xNew THEN
    FOR uiI := UINT#0 TO UINT#119 DO aSeen[uiI] := aFrame[uiI]; END_FOR;
    FOR uiI := UINT#0 TO UINT#117 DO
        aFrameBytes[uiI * UINT#2] := WORD_TO_BYTE(SHR(aFrame[uiI], 8));
        aFrameBytes[uiI * UINT#2 + UINT#1] := WORD_TO_BYTE(aFrame[uiI] AND WORD#255);
    END_FOR;
    FOR uiI := UINT#0 TO UINT#95 DO
        aPayload[uiI * UINT#2] := WORD_TO_BYTE(SHR(aFrame[uiI + UINT#20], 8));
        aPayload[uiI * UINT#2 + UINT#1] := WORD_TO_BYTE(aFrame[uiI + UINT#20] AND WORD#255);
    END_FOR;
    uiOp := WORD_TO_UINT(aFrame[2]);
    udiSeq := SHL(WORD_TO_UDINT(aFrame[3]), 16) OR WORD_TO_UDINT(aFrame[4]);
    udiSession := SHL(WORD_TO_UDINT(aFrame[5]), 16) OR WORD_TO_UDINT(aFrame[6]);
    udiBoot := SHL(WORD_TO_UDINT(aFrame[7]), 16) OR WORD_TO_UDINT(aFrame[8]);
    udiFrameSize := SHL(WORD_TO_UDINT(aFrame[9]), 16) OR WORD_TO_UDINT(aFrame[10]);
    udiOffset := SHL(WORD_TO_UDINT(aFrame[11]), 16) OR WORD_TO_UDINT(aFrame[12]);
    uiLength := WORD_TO_UINT(aFrame[13]);
    udiFileCrc := SHL(WORD_TO_UDINT(aFrame[14]), 16) OR WORD_TO_UDINT(aFrame[15]);
    udiFrameCrc := F_FileCrc32(ADR(aFrameBytes), UINT#236, UDINT#16#FFFFFFFF) XOR UDINT#16#FFFFFFFF;
    wRequestError := WORD#0;
    xAccept := FALSE;
    IF (aFrame[0] <> WORD#16#F7B1) OR (aFrame[1] <> WORD#1)
        OR (aFrame[19] <> WORD#0) OR (aFrame[116] <> WORD#0) OR (aFrame[117] <> WORD#0)
        OR (uiLength > UINT#192) OR (udiSeq = UDINT#0) OR (udiSession = UDINT#0) THEN
        wRequestError := WORD#16#E001;
    ELSIF udiFrameCrc <> (SHL(WORD_TO_UDINT(aFrame[118]), 16) OR WORD_TO_UDINT(aFrame[119])) THEN
        wRequestError := WORD#16#E002;
    ELSIF udiBoot <> GVL_FileBridgeRetain.udiBootCounter THEN
        wRequestError := WORD#16#E003;
    ELSIF (udiSession = udiOwner) AND (udiSeq = udiAck) THEN
        xSame := TRUE;
        FOR uiI := UINT#0 TO UINT#119 DO
            IF aAccepted[uiI] <> aFrame[uiI] THEN xSame := FALSE; END_IF;
        END_FOR;
        IF NOT xSame THEN wRequestError := WORD#16#E004; END_IF;
        (* Exact replay: existing ACK/status only; NEVER repeat file/FTP operations. *)
    ELSE
        IF (uiOp = UINT#1) AND ((uiState = UINT#0) OR (uiState = UINT#400)) THEN
            IF (udiSeq <> UDINT#1) OR NOT xClean THEN wRequestError := WORD#16#E005; END_IF;
        ELSIF udiSession <> udiOwner THEN
            wRequestError := WORD#16#E006;
        ELSIF (udiSeq <= udiAck) OR (udiAck = UDINT#16#FFFFFFFF) THEN
            wRequestError := WORD#16#E005;
        ELSIF (uiOp <> UINT#4) AND (uiOp <> UINT#6) AND (udiSeq <> udiAck + UDINT#1) THEN
            wRequestError := WORD#16#E005;
        END_IF;
        IF NOT GVL_FileBridge.xFileTransferPermit AND (uiOp <> UINT#4) AND (uiOp <> UINT#6) THEN
            wRequestError := WORD#16#E007;
        END_IF;
        IF wRequestError = WORD#0 THEN
            CASE uiOp OF
                UINT#1: (* START file; first file also creates project session. *)
                    sNewProject := '';
                    sNewFile := '';
                    uiField := UINT#0;
                    uiPos := UINT#0;
                    xNamesOk := (uiLength >= UINT#2) AND (uiLength <= UINT#98);
                    IF xNamesOk THEN
                        FOR uiI := UINT#0 TO uiLength - UINT#1 DO
                            IF uiField = UINT#0 THEN pName := ADR(sNewProject);
                            ELSE pName := ADR(sNewFile); END_IF;
                            IF aPayload[uiI] = BYTE#0 THEN
                                IF uiPos = UINT#0 THEN xNamesOk := FALSE; END_IF;
                                uiField := uiField + UINT#1;
                                uiPos := UINT#0;
                            ELSIF (uiField > UINT#1) OR (uiPos >= UINT#48) THEN
                                xNamesOk := FALSE;
                            ELSE
                                pName[uiPos] := aPayload[uiI];
                                uiPos := uiPos + UINT#1;
                                pName[uiPos] := BYTE#0;
                            END_IF;
                        END_FOR;
                    END_IF;
                    xNamesOk := xNamesOk AND (uiField = UINT#2) AND (uiPos = UINT#0)
                        AND F_FileNameValid(sNewProject, TRUE) AND F_FileNameValid(sNewFile, FALSE);
                    uiCount := WORD_TO_UINT(aFrame[16]);
                    uiIndex := WORD_TO_UINT(aFrame[17]);
                    IF NOT GVL_FileBridge.xFileTransferPermit THEN
                        wRequestError := WORD#16#E007;
                    ELSIF NOT xNamesOk OR (aFrame[18] > WORD#2) THEN
                        wRequestError := WORD#16#E008;
                    ELSIF (aFrame[18] = WORD#2) AND (NOT xFixedConfig
                        OR NOT GVL_FileBridge.xFixedIdle OR (sNewProject <> GVL_FileBridge.sFixedProject)
                        OR (uiCount <> UINT#7) OR NOT F_FixedFileValid(sNewFile)) THEN
                        wRequestError := WORD#16#E015;
                    ELSIF (aFrame[18] <> WORD#2) AND (sNewProject = GVL_FileBridge.sFixedProject) THEN
                        wRequestError := WORD#16#E015;
                    ELSIF (udiFrameSize > UDINT#1048576)
                        OR (uiCount = UINT#0) OR (uiCount > UINT#32) OR (udiOffset <> UDINT#0) THEN
                        wRequestError := WORD#16#E009;
                    ELSIF (aFrame[18] = WORD#1) AND (RIGHT(sNewFile, 4) = '.txt') THEN
                        wRequestError := WORD#16#E008;
                    ELSIF (uiState = UINT#0) OR (uiState = UINT#400) THEN
                        IF (uiIndex <> UINT#1) OR (udiSeq <> UDINT#1) THEN
                            wRequestError := WORD#16#E00A;
                        ELSE
                            udiOwner := udiSession;
                            uiVerified := UINT#0;
                            udiTotalSize := UDINT#0;
                            uiExpectedFiles := uiCount;
                            uiMode := WORD_TO_UINT(aFrame[18]);
                            sProject := sNewProject;
                            IF uiMode = UINT#2 THEN
                                GVL_FileBridge.xFixedReady := FALSE;
                                GVL_FileBridge.xFixedUpdateBusy := TRUE;
                                uiSessionCapture := GVL_FileBridge.uiFixedCapture;
                                uiSessionPath := GVL_FileBridge.uiFixedPath;
                                uiSessionReturn := GVL_FileBridge.uiFixedReturn;
                            END_IF;
                            xAccept := TRUE;
                        END_IF;
                    ELSIF (uiState <> UINT#200) OR (sNewProject <> sProject)
                        OR (uiIndex <> uiVerified + UINT#1) OR (uiIndex > uiExpectedFiles)
                        OR (uiCount <> uiExpectedFiles) OR (aFrame[18] <> UINT_TO_WORD(uiMode)) THEN
                        wRequestError := WORD#16#E00A;
                    ELSE
                        xAccept := TRUE;
                        FOR uiI := UINT#0 TO uiVerified - UINT#1 DO
                            IF aNames[uiI] = sNewFile THEN
                                xAccept := FALSE;
                                wRequestError := WORD#16#E00B;
                            END_IF;
                        END_FOR;
                    END_IF;
                    IF xAccept THEN
                        IF udiTotalSize + udiFrameSize > UDINT#5242880 THEN
                            xAccept := FALSE;
                            wRequestError := WORD#16#E009;
                        ELSE
                            sFile := sNewFile;
                            udiSize := udiFrameSize;
                            udiExpectedCrc := udiFileCrc;
                            udiRunningCrc := UDINT#16#FFFFFFFF;
                            udiReceived := UDINT#0;
                            uiOrdinal := uiIndex;
                            uiState := UINT#100;
                            wError := WORD#0;
                            xFileVerified := FALSE;
                        END_IF;
                    END_IF;
                UINT#2: (* CHUNK; sequential, no writes while FTP owns buffer. *)
                    IF (uiState <> UINT#100) OR (uiLength = UINT#0)
                        OR (udiOffset <> udiReceived) OR (udiOffset + UINT_TO_UDINT(uiLength) > udiSize) THEN
                        wRequestError := WORD#16#E00C;
                    ELSE
                        FOR uiI := UINT#0 TO uiLength - UINT#1 DO
                            GVL_FileBridge.aBuffer[udiReceived + UINT_TO_UDINT(uiI)] := aPayload[uiI];
                        END_FOR;
                        udiRunningCrc := F_FileCrc32(ADR(aPayload), uiLength, udiRunningCrc);
                        udiReceived := udiReceived + UINT_TO_UDINT(uiLength);
                        xAccept := TRUE;
                    END_IF;
                UINT#3: (* DEPLOY only complete, CRC-checked RAM image. *)
                    IF (uiState <> UINT#100) OR (udiReceived <> udiSize) OR (uiLength <> UINT#0) THEN
                        wRequestError := WORD#16#E00D;
                    ELSIF (udiRunningCrc XOR UDINT#16#FFFFFFFF) <> udiExpectedCrc THEN
                        wRequestError := WORD#16#E00E;
                        wError := wRequestError;
                        uiState := UINT#900;
                    ELSIF NOT GVL_FileBridge.xFileTransferPermit THEN
                        wRequestError := WORD#16#E007;
                    ELSE
                        uiState := UINT#300;
                        xAccept := TRUE;
                    END_IF;
                UINT#4: (* ABORT; cleanup cannot be skipped or rearmed remotely. *)
                    IF (uiState = UINT#300) OR (uiState = UINT#310) THEN
                        uiState := UINT#310;
                    ELSE
                        uiState := UINT#900;
                    END_IF;
                    wError := WORD#16#E010;
                    xAccept := TRUE;
                UINT#5: (* FINISH: all files individually uploaded AND read back. *)
                    IF (uiState <> UINT#200) OR (uiVerified <> uiExpectedFiles) THEN
                        wRequestError := WORD#16#E00F;
                    ELSIF (uiMode = UINT#2) AND (NOT xFixedConfig OR NOT GVL_FileBridge.xFixedIdle
                        OR (sProject <> GVL_FileBridge.sFixedProject)
                        OR (uiSessionCapture <> GVL_FileBridge.uiFixedCapture)
                        OR (uiSessionPath <> GVL_FileBridge.uiFixedPath)
                        OR (uiSessionReturn <> GVL_FileBridge.uiFixedReturn)) THEN
                        wRequestError := WORD#16#E015;
                    ELSE
                        xPairsOk := TRUE;
                        IF (uiMode = UINT#1) OR (uiMode = UINT#2) THEN
                            xGlobal := FALSE;
                            uiPrograms := UINT#0;
                            FOR uiI := UINT#0 TO uiVerified - UINT#1 DO
                                IF aNames[uiI] = '_project.srd' THEN xGlobal := TRUE; END_IF;
                                IF RIGHT(aNames[uiI], 4) = '.srp' THEN
                                    uiPrograms := uiPrograms + UINT#1;
                                    sPair := CONCAT(LEFT(aNames[uiI], LEN(aNames[uiI]) - 1), 'd');
                                    xFound := FALSE;
                                    FOR uiJ := UINT#0 TO uiVerified - UINT#1 DO
                                        IF aNames[uiJ] = sPair THEN xFound := TRUE; END_IF;
                                    END_FOR;
                                    IF NOT xFound THEN xPairsOk := FALSE; END_IF;
                                END_IF;
                            END_FOR;
                            xPairsOk := xPairsOk AND xGlobal AND (uiPrograms > UINT#0);
                        END_IF;
                        IF xPairsOk THEN
                            uiState := UINT#400; xAccept := TRUE;
                            IF uiMode = UINT#2 THEN
                                GVL_FileBridge.xFixedReady := TRUE;
                                sReadyProject := GVL_FileBridge.sFixedProject;
                                uiReadyCapture := GVL_FileBridge.uiFixedCapture;
                                uiReadyPath := GVL_FileBridge.uiFixedPath;
                                uiReadyReturn := GVL_FileBridge.uiFixedReturn;
                            END_IF;
                        ELSE wRequestError := WORD#16#E012; END_IF;
                    END_IF;
                UINT#6: (* RELEASE only after all handles are known closed. *)
                    IF xClean AND ((uiState = UINT#400) OR (uiState = UINT#900)) THEN
                        uiState := UINT#0;
                        xAccept := TRUE;
                    ELSE wRequestError := WORD#16#E013; END_IF;
            ELSE
                wRequestError := WORD#16#E001;
            END_CASE;
        END_IF;
        IF xAccept THEN
            udiAck := udiSeq;
            uiAckOp := uiOp;
            FOR uiI := UINT#0 TO UINT#119 DO aAccepted[uiI] := aFrame[uiI]; END_FOR;
        END_IF;
    END_IF;
    IF wRequestError <> WORD#0 THEN
        wReject := wRequestError;
        udiRejectSeq := udiSeq;
        udiRejectOwner := udiSession;
    END_IF;
END_IF;

IF xActive AND (fbLease.Q OR NOT GVL_FileBridge.xFileTransferPermit
    OR ((uiMode = UINT#2) AND (NOT xFixedConfig OR NOT GVL_FileBridge.xFixedIdle
        OR (sProject <> GVL_FileBridge.sFixedProject)
        OR (uiSessionCapture <> GVL_FileBridge.uiFixedCapture)
        OR (uiSessionPath <> GVL_FileBridge.uiFixedPath)
        OR (uiSessionReturn <> GVL_FileBridge.uiFixedReturn)))) THEN
    IF fbLease.Q THEN wError := WORD#16#E011;
    ELSE wError := WORD#16#E007; END_IF;
    IF (uiState = UINT#300) OR (uiState = UINT#310) THEN uiState := UINT#310;
    ELSIF uiState <> UINT#400 THEN uiState := UINT#900; END_IF;
END_IF;

IF ((uiState = UINT#300) OR (uiState = UINT#310)) AND xFtpStarted AND fbFtp.xDone THEN
    xFtpStarted := FALSE;
    IF (uiState = UINT#300) AND fbFtp.xTestPassed THEN
        aNames[uiVerified] := sFile;
        uiVerified := uiVerified + UINT#1;
        udiTotalSize := udiTotalSize + udiSize;
        xFileVerified := TRUE;
        uiState := UINT#200;
    ELSE
        IF wError = WORD#0 THEN wError := WORD#16#E014; END_IF;
        IF fbFtp.xControlOwned OR fbFtp.xDataOwned THEN uiState := UINT#910;
        ELSE uiState := UINT#900; END_IF;
    END_IF;
END_IF;
IF (uiState = UINT#300) OR (uiState = UINT#310) THEN xFtpStarted := TRUE; END_IF;
fbFtp(xStart := (uiState = UINT#300) OR (uiState = UINT#310),
    xAbort := uiState = UINT#310, pBuffer := ADR(GVL_FileBridge.aBuffer),
    udiSize := udiSize, sProject := sProject, sFile := sFile,
    xCreateProject := uiVerified = UINT#0,
    xReplaceFixed := uiMode = UINT#2,
    sUser := GVL_FileBridge.sFtpUser, sPassword := GVL_FileBridge.sFtpPassword);

(* Coherent FC03 status: matching EVEN snapshot head/tail required by PC. *)
IF uiSnapshot >= UINT#65534 THEN uiSnapshot := UINT#0;
ELSE uiSnapshot := uiSnapshot + UINT#2; END_IF;
GVL_FileBridge.aStatus[38] := UINT_TO_WORD(uiSnapshot + UINT#1);
wFlags := WORD#0;
IF GVL_FileBridge.xFileTransferPermit THEN wFlags := wFlags OR WORD#1; END_IF;
IF xClean THEN wFlags := wFlags OR WORD#2; END_IF;
IF xFileVerified THEN wFlags := wFlags OR WORD#4; END_IF;
IF uiState = UINT#400 THEN wFlags := wFlags OR WORD#8; END_IF;
IF (uiState = UINT#300) OR (uiState = UINT#310) THEN wFlags := wFlags OR WORD#16; END_IF;
GVL_FileBridge.aStatus[0] := WORD#16#F7B2;
GVL_FileBridge.aStatus[1] := WORD#1;
GVL_FileBridge.aStatus[2] := UINT_TO_WORD(uiState);
GVL_FileBridge.aStatus[3] := wError;
GVL_FileBridge.aStatus[4] := UDINT_TO_WORD(SHR(udiAck, 16));
GVL_FileBridge.aStatus[5] := UDINT_TO_WORD(udiAck);
GVL_FileBridge.aStatus[6] := UINT_TO_WORD(uiAckOp);
GVL_FileBridge.aStatus[7] := wFlags;
GVL_FileBridge.aStatus[8] := UDINT_TO_WORD(SHR(udiOwner, 16));
GVL_FileBridge.aStatus[9] := UDINT_TO_WORD(udiOwner);
GVL_FileBridge.aStatus[10] := UDINT_TO_WORD(SHR(GVL_FileBridgeRetain.udiBootCounter, 16));
GVL_FileBridge.aStatus[11] := UDINT_TO_WORD(GVL_FileBridgeRetain.udiBootCounter);
GVL_FileBridge.aStatus[12] := UDINT_TO_WORD(SHR(udiReceived, 16));
GVL_FileBridge.aStatus[13] := UDINT_TO_WORD(udiReceived);
GVL_FileBridge.aStatus[14] := UDINT_TO_WORD(SHR(udiSize, 16));
GVL_FileBridge.aStatus[15] := UDINT_TO_WORD(udiSize);
GVL_FileBridge.aStatus[16] := UDINT_TO_WORD(SHR(udiRunningCrc XOR UDINT#16#FFFFFFFF, 16));
GVL_FileBridge.aStatus[17] := UDINT_TO_WORD(udiRunningCrc XOR UDINT#16#FFFFFFFF);
GVL_FileBridge.aStatus[18] := UDINT_TO_WORD(SHR(udiExpectedCrc, 16));
GVL_FileBridge.aStatus[19] := UDINT_TO_WORD(udiExpectedCrc);
GVL_FileBridge.aStatus[20] := UINT_TO_WORD(uiVerified);
GVL_FileBridge.aStatus[21] := UINT_TO_WORD(uiExpectedFiles);
GVL_FileBridge.aStatus[22] := UINT_TO_WORD(uiOrdinal);
GVL_FileBridge.aStatus[23] := UINT_TO_WORD(fbFtp.uiStep);
GVL_FileBridge.aStatus[24] := UINT_TO_WORD(fbFtp.uiReplyCode);
GVL_FileBridge.aStatus[25] := fbFtp.wErrorID;
GVL_FileBridge.aStatus[26] := UINT_TO_WORD(fbFtp.uiErrorStage);
GVL_FileBridge.aStatus[27] := UDINT_TO_WORD(SHR(fbFtp.udiUploadedBytes, 16));
GVL_FileBridge.aStatus[28] := UDINT_TO_WORD(fbFtp.udiUploadedBytes);
GVL_FileBridge.aStatus[29] := UDINT_TO_WORD(SHR(fbFtp.udiReadbackBytes, 16));
GVL_FileBridge.aStatus[30] := UDINT_TO_WORD(fbFtp.udiReadbackBytes);
GVL_FileBridge.aStatus[31] := wReject;
GVL_FileBridge.aStatus[32] := UDINT_TO_WORD(SHR(udiRejectSeq, 16));
GVL_FileBridge.aStatus[33] := UDINT_TO_WORD(udiRejectSeq);
GVL_FileBridge.aStatus[34] := UDINT_TO_WORD(SHR(udiRejectOwner, 16));
GVL_FileBridge.aStatus[35] := UDINT_TO_WORD(udiRejectOwner);
GVL_FileBridge.aStatus[36] := wHeartbeatOld;
GVL_FileBridge.aStatus[37] := WORD#32;
GVL_FileBridge.aStatus[39] := WORD#16;
GVL_FileBridge.aStatus[40] := WORD#0;
GVL_FileBridge.aStatus[41] := WORD#192;
GVL_FileBridge.aStatus[42] := fbFtp.wDataCloseErrorID;
GVL_FileBridge.aStatus[43] := fbFtp.wControlCloseErrorID;
GVL_FileBridge.aStatus[44] := UINT_TO_WORD(uiMode);
GVL_FileBridge.aStatus[45] := UINT_TO_WORD(fbFtp.uiUploadCompleteCode);
GVL_FileBridge.aStatus[46] := UINT_TO_WORD(fbFtp.uiDownloadCompleteCode);
GVL_FileBridge.aStatus[47] := WORD#3; (* bit0 empty files; bit1 guarded fixed-project replacement *)
GVL_FileBridge.aStatus[48] := WORD#16#0102;
FOR uiI := UINT#49 TO UINT#62 DO GVL_FileBridge.aStatus[uiI] := WORD#0; END_FOR;
IF xFixedConfig THEN GVL_FileBridge.aStatus[49] := WORD#1; END_IF;
GVL_FileBridge.xFixedUpdateBusy := (uiMode = UINT#2) AND ((uiState = UINT#100)
    OR (uiState = UINT#200) OR (uiState = UINT#300) OR (uiState = UINT#310) OR (uiState = UINT#910));
IF GVL_FileBridge.xFixedUpdateBusy THEN GVL_FileBridge.aStatus[50] := WORD#1; END_IF;
IF GVL_FileBridge.xFixedReady THEN GVL_FileBridge.aStatus[51] := WORD#1; END_IF;
GVL_FileBridge.aStatus[52] := UINT_TO_WORD(GVL_FileBridge.uiFixedCapture);
GVL_FileBridge.aStatus[53] := UINT_TO_WORD(GVL_FileBridge.uiFixedPath);
GVL_FileBridge.aStatus[54] := UINT_TO_WORD(GVL_FileBridge.uiFixedReturn);
GVL_FileBridge.aStatus[55] := UDINT_TO_WORD(SHR(udiFixedProjectCrc, 16));
GVL_FileBridge.aStatus[56] := UDINT_TO_WORD(udiFixedProjectCrc);
IF GVL_FileBridge.xFixedIdle THEN GVL_FileBridge.aStatus[59] := WORD#1; END_IF;
GVL_FileBridge.aStatus[63] := UINT_TO_WORD(uiSnapshot);
GVL_FileBridge.aStatus[38] := UINT_TO_WORD(uiSnapshot);
END_PROGRAM

(* ---- PRG_RobotBridge.st ---- *)
PROGRAM PRG_RobotBridge
VAR
    xFirstScan : BOOL := TRUE;
    i : INT;
    xSame : BOOL;
    xNewFrame : BOOL;
    uiStable : UINT;
    aPrevious : ARRAY[0..14] OF WORD;
    aConsumed : ARRAY[0..14] OF WORD;
    aFrame : ARRAY[0..15] OF WORD;
    udiRequest : UDINT;
    udiRequestHost : UDINT;
    udiExpectedBoot : UDINT;
    udiOwner : UDINT;
    udiLastSeq : UDINT;
    udiAckSeq : UDINT;
    udiRejectedSeq : UDINT;
    udiInterruptedSeq : UDINT;
    wAckCmd : WORD;
    wAckResult : WORD;
    wAckError : WORD;
    wReject : WORD;
    wLastReject : WORD;
    wCmd : WORD;
    wParam : WORD;
    wPlcHb : WORD;
    wLastHostHb : WORD;
    xHostHbEdge : BOOL;
    xHb : BOOL;
    xLastHb : BOOL;
    xHbEdge : BOOL;
    uiHbEdges : UINT;
    wHbCount : WORD;
    fbRobotTimeout : TON;
    fbHostTimeout : TON;
    uiStep : UINT;
    wPulse : WORD;
    uiSelectedProgram : UINT;
    xCoordinates : BOOL;
    xLoadSent : BOOL;
    xHasControlledRobot : BOOL;
    xNewAction : BOOL;
    xConfirmed : BOOL;
    xRunningSeen : BOOL;
    xTerminalStop : BOOL;
    wCancelReason : WORD;
    wFlags : WORD;
    fbLowBefore : TON;
    fbPulse : TON;
    fbLowAfter : TON;
    fbActionTimeout : TON;
END_VAR

GVL_RobotBridge.uiFixedJobGuardVersion := UINT#120;

// ----- Startup: ignore retained/stale command frames -----
IF xFirstScan THEN
    IF GVL_RobotBridgeRetain.udiBootCounter = UDINT#4294967295 THEN
        GVL_RobotBridgeRetain.udiBootCounter := UDINT#1;
    ELSE
        GVL_RobotBridgeRetain.udiBootCounter :=
            GVL_RobotBridgeRetain.udiBootCounter + UDINT#1;
    END_IF;
    FOR i := 0 TO 14 DO
        aPrevious[i] := GVL_RobotBridge.aHostCmd[i];
        aConsumed[i] := GVL_RobotBridge.aHostCmd[i];
    END_FOR;
    xLastHb := (GVL_RobotBridge.aRobotRx[0] AND WORD#16#0200) <> WORD#0;
    wLastHostHb := GVL_RobotBridge.aHostCmd[15];
    xFirstScan := FALSE;
END_IF;

// ----- STEP status: DO33..48 in the first input register -----
GVL_RobotBridge.xRobotRunning := (GVL_RobotBridge.aRobotRx[0] AND WORD#16#0001) <> WORD#0;
GVL_RobotBridge.xRobotAlarm := (GVL_RobotBridge.aRobotRx[0] AND WORD#16#0002) <> WORD#0;
GVL_RobotBridge.xRobotEnabled := (GVL_RobotBridge.aRobotRx[0] AND WORD#16#0004) <> WORD#0;
GVL_RobotBridge.xRobotPaused := (GVL_RobotBridge.aRobotRx[0] AND WORD#16#0008) <> WORD#0;
GVL_RobotBridge.xRobotStopped := (GVL_RobotBridge.aRobotRx[0] AND WORD#16#0010) <> WORD#0;
GVL_RobotBridge.xRobotExternalAuto := (GVL_RobotBridge.aRobotRx[0] AND WORD#16#0080) <> WORD#0;
GVL_RobotBridge.xRobotEmergency := (GVL_RobotBridge.aRobotRx[0] AND WORD#16#0100) <> WORD#0;
IF NOT GVL_RobotBridge.xRobotExternalAuto OR GVL_RobotBridge.xRobotAlarm
   OR GVL_RobotBridge.xRobotEmergency OR GVL_FileBridge.xFixedUpdateBusy THEN
    GVL_RobotBridge.xLoadOperatorConfirmed := FALSE;
END_IF;
IF GVL_FileBridge.xFixedUpdateBusy THEN xLoadSent := FALSE; END_IF;
xTerminalStop := GVL_RobotBridge.xRobotStopped
    AND NOT GVL_RobotBridge.xRobotRunning AND NOT GVL_RobotBridge.xRobotPaused;
xHb := (GVL_RobotBridge.aRobotRx[0] AND WORD#16#0200) <> WORD#0;
xHbEdge := xHb <> xLastHb;
xLastHb := xHb;
fbRobotTimeout(IN := NOT xHbEdge, PT := T#4s);
IF fbRobotTimeout.Q OR GVL_RobotBridge.xNativeModbusError THEN
    uiHbEdges := UINT#0;
ELSIF xHbEdge AND (uiHbEdges < UINT#2) THEN
    uiHbEdges := uiHbEdges + UINT#1;
END_IF;
IF xHbEdge THEN
    IF wHbCount = WORD#16#FFFF THEN wHbCount := WORD#0;
    ELSE wHbCount := UINT_TO_WORD(WORD_TO_UINT(wHbCount) + UINT#1); END_IF;
END_IF;
GVL_RobotBridge.xRobotLinkOK := (uiHbEdges >= UINT#2)
    AND NOT fbRobotTimeout.Q AND NOT GVL_RobotBridge.xNativeModbusError;

// ----- Only the registered owner can refresh its heartbeat -----
udiRequestHost := SHL(WORD_TO_UDINT(GVL_RobotBridge.aHostCmd[6]), 16)
    OR WORD_TO_UDINT(GVL_RobotBridge.aHostCmd[7]);
udiExpectedBoot := SHL(WORD_TO_UDINT(GVL_RobotBridge.aHostCmd[8]), 16)
    OR WORD_TO_UDINT(GVL_RobotBridge.aHostCmd[9]);
xHostHbEdge := GVL_RobotBridge.xHostRegistered
    AND (GVL_RobotBridge.aHostCmd[0] = WORD#2)
    AND (udiRequestHost = udiOwner)
    AND (udiExpectedBoot = GVL_RobotBridgeRetain.udiBootCounter)
    AND (GVL_RobotBridge.aHostCmd[15] <> wLastHostHb);
IF xHostHbEdge THEN wLastHostHb := GVL_RobotBridge.aHostCmd[15]; END_IF;
fbHostTimeout(IN := GVL_RobotBridge.xHostRegistered AND NOT xHostHbEdge, PT := T#3s);
GVL_RobotBridge.xHostAlive := GVL_RobotBridge.xHostRegistered AND NOT fbHostTimeout.Q;
IF fbHostTimeout.Q THEN
    GVL_RobotBridge.xHostRegistered := FALSE;
    GVL_RobotBridge.xHostAlive := FALSE;
    udiOwner := UDINT#0;
END_IF;

// ----- Ordinary stop interlock; never represents a safety-rated stop -----
wCancelReason := WORD#0;
IF NOT GVL_RobotBridge.xCommissioned OR NOT GVL_RobotBridge.xGdiProgramMappingConfirmed THEN
    wCancelReason := WORD#13;
ELSIF NOT GVL_RobotBridge.xRemotePermit THEN wCancelReason := WORD#6;
ELSIF NOT GVL_RobotBridge.xRobotLinkOK THEN wCancelReason := WORD#7;
ELSIF NOT GVL_RobotBridge.xHostAlive THEN wCancelReason := WORD#11;
ELSIF GVL_RobotBridge.xRobotEmergency THEN wCancelReason := WORD#12;
ELSIF GVL_RobotBridge.xRobotAlarm AND (wAckCmd <> WORD#8)
      AND (wAckCmd <> WORD#7) THEN wCancelReason := WORD#12;
END_IF;
IF xHasControlledRobot AND (wCancelReason <> WORD#0) THEN
    GVL_RobotBridge.xStopInterlock := TRUE;
    GVL_RobotBridge.xLoadOperatorConfirmed := FALSE;
    IF (uiStep <> UINT#0) AND NOT ((wAckCmd = WORD#7)
       AND GVL_RobotBridge.xCommissioned AND GVL_RobotBridge.xRobotLinkOK
       AND GVL_RobotBridge.xHostAlive) THEN
        uiStep := UINT#0;
        wAckResult := WORD#6;
        wAckError := wCancelReason;
        wPulse := WORD#0;
    END_IF;
END_IF;

// ----- Stable command snapshot, heartbeat excluded -----
FOR i := 0 TO 15 DO aFrame[i] := GVL_RobotBridge.aHostCmd[i]; END_FOR;
xSame := TRUE;
FOR i := 0 TO 14 DO
    IF aFrame[i] <> aPrevious[i] THEN xSame := FALSE; END_IF;
    aPrevious[i] := aFrame[i];
END_FOR;
IF xSame THEN
    IF uiStable < UINT#2 THEN uiStable := uiStable + UINT#1; END_IF;
ELSE uiStable := UINT#0;
END_IF;
xNewFrame := FALSE;
IF uiStable >= UINT#2 THEN
    FOR i := 0 TO 14 DO
        IF aFrame[i] <> aConsumed[i] THEN xNewFrame := TRUE; END_IF;
    END_FOR;
END_IF;
xNewAction := FALSE;
IF xNewFrame THEN
    FOR i := 0 TO 14 DO aConsumed[i] := aFrame[i]; END_FOR;
    wCmd := aFrame[1];
    wParam := aFrame[4];
    udiRequest := SHL(WORD_TO_UDINT(aFrame[2]), 16) OR WORD_TO_UDINT(aFrame[3]);
    udiRequestHost := SHL(WORD_TO_UDINT(aFrame[6]), 16) OR WORD_TO_UDINT(aFrame[7]);
    udiExpectedBoot := SHL(WORD_TO_UDINT(aFrame[8]), 16) OR WORD_TO_UDINT(aFrame[9]);
    wReject := WORD#0;
    IF aFrame[0] <> WORD#2 THEN wReject := WORD#1;
    ELSIF (udiRequest = UDINT#0) OR (udiRequestHost = UDINT#0) THEN wReject := WORD#8;
    ELSIF udiExpectedBoot <> GVL_RobotBridgeRetain.udiBootCounter THEN wReject := WORD#3;
    ELSIF (wCmd <> WORD#4) AND (wCmd <> WORD#10) AND (wCmd <> WORD#12)
          AND (wParam <> WORD#0) THEN wReject := WORD#8;
    ELSE
        FOR i := 5 TO 14 DO
            IF ((i = 5) OR (i >= 10)) AND (aFrame[i] <> WORD#0) THEN wReject := WORD#14; END_IF;
        END_FOR;
    END_IF;

    IF wReject = WORD#0 THEN
        IF wCmd = WORD#1 THEN
            IF (uiStep <> UINT#0) OR (GVL_RobotBridge.xHostRegistered AND (udiOwner <> udiRequestHost)) THEN
                wReject := WORD#2;
            ELSIF GVL_RobotBridge.xHostRegistered AND (udiRequest <= udiLastSeq) THEN
                wReject := WORD#4;
            ELSE
                udiOwner := udiRequestHost;
                udiLastSeq := udiRequest;
                GVL_RobotBridge.xHostRegistered := TRUE;
                GVL_RobotBridge.xHostAlive := TRUE;
                wLastHostHb := aFrame[15];
                udiAckSeq := udiRequest; wAckCmd := wCmd;
                wAckResult := WORD#2; wAckError := WORD#0;
            END_IF;
        ELSIF NOT GVL_RobotBridge.xHostRegistered OR (udiOwner <> udiRequestHost) THEN
            wReject := WORD#2;
        ELSIF udiRequest <= udiLastSeq THEN wReject := WORD#4;
        ELSE
            udiLastSeq := udiRequest;
            IF (uiStep <> UINT#0) AND (wCmd <> WORD#7) THEN wReject := WORD#5;
            ELSE
                // STOP can preempt the one active request; preserve its sequence.
                IF uiStep <> UINT#0 THEN
                    udiInterruptedSeq := udiAckSeq;
                    uiStep := UINT#0;
                    wPulse := WORD#0;
                END_IF;
                udiAckSeq := udiRequest; wAckCmd := wCmd;
                wAckResult := WORD#2; wAckError := WORD#0;
                IF (wCmd >= WORD#2) AND (wCmd <= WORD#8) THEN
                    IF NOT GVL_RobotBridge.xCommissioned THEN wReject := WORD#13;
                    ELSIF NOT GVL_RobotBridge.xGdiProgramMappingConfirmed
                          AND (wCmd <> WORD#3) AND (wCmd <> WORD#7) AND (wCmd <> WORD#8) THEN
                        wReject := WORD#13;
                    ELSIF NOT GVL_RobotBridge.xRobotLinkOK THEN wReject := WORD#7;
                    ELSIF (wCmd <> WORD#7) AND NOT GVL_RobotBridge.xRemotePermit THEN wReject := WORD#6;
                    ELSIF (wCmd <> WORD#7) AND GVL_RobotBridge.xStopInterlock THEN wReject := WORD#15;
                    ELSIF NOT GVL_RobotBridge.xHostAlive THEN wReject := WORD#11;
                    ELSIF GVL_FileBridge.xFixedUpdateBusy AND ((wCmd = WORD#2) OR (wCmd = WORD#4) OR (wCmd = WORD#5)) THEN
                        wReject := WORD#9;
                    END_IF;
                    IF wReject = WORD#0 THEN
                        wPulse := WORD#0;
                        CASE WORD_TO_UINT(wCmd) OF
                        2: // Enable is a toggle input: pulse ONLY when currently disabled.
                            IF NOT xTerminalStop OR NOT GVL_RobotBridge.xRobotExternalAuto
                               OR GVL_RobotBridge.xRobotAlarm OR GVL_RobotBridge.xRobotEmergency THEN
                                wReject := WORD#9;
                            ELSIF NOT GVL_RobotBridge.xRobotEnabled THEN wPulse := WORD#16#0010; END_IF;
                        3: // Disable: same toggle input, only while stopped.
                            IF NOT xTerminalStop THEN wReject := WORD#9;
                            ELSIF GVL_RobotBridge.xRobotEnabled THEN wPulse := WORD#16#0010; END_IF;
                        4: // GDI DI49..56: unsigned binary program number 1..255.
                            IF (wParam < WORD#1) OR (wParam > WORD#255) THEN wReject := WORD#8;
                            ELSIF GVL_FileBridge.xFixedMappingConfirmed AND NOT GVL_FileBridge.xFixedReady
                                AND ((wParam = UINT_TO_WORD(GVL_FileBridge.uiFixedCapture))
                                    OR (wParam = UINT_TO_WORD(GVL_FileBridge.uiFixedPath))
                                    OR (wParam = UINT_TO_WORD(GVL_FileBridge.uiFixedReturn))) THEN wReject := WORD#9;
                            ELSIF NOT xTerminalStop OR NOT GVL_RobotBridge.xRobotExternalAuto
                                  OR GVL_RobotBridge.xRobotAlarm OR GVL_RobotBridge.xRobotEmergency THEN
                                wReject := WORD#9;
                            ELSE
                                uiSelectedProgram := WORD_TO_UINT(wParam);
                                xLoadSent := FALSE;
                                GVL_RobotBridge.xLoadOperatorConfirmed := FALSE;
                                wPulse := WORD#16#0020;
                            END_IF;
                        5: // Run/resume requires enable and an explicit confirmed loaded program.
                            IF GVL_FileBridge.xFixedMappingConfirmed AND NOT GVL_FileBridge.xFixedReady
                                AND ((uiSelectedProgram = GVL_FileBridge.uiFixedCapture)
                                    OR (uiSelectedProgram = GVL_FileBridge.uiFixedPath)
                                    OR (uiSelectedProgram = GVL_FileBridge.uiFixedReturn)) THEN wReject := WORD#9;
                            ELSIF NOT GVL_RobotBridge.xRobotExternalAuto OR NOT GVL_RobotBridge.xRobotEnabled
                               OR GVL_RobotBridge.xRobotAlarm OR GVL_RobotBridge.xRobotEmergency
                               OR NOT GVL_RobotBridge.xLoadOperatorConfirmed
                               OR NOT (xTerminalStop OR GVL_RobotBridge.xRobotPaused) THEN wReject := WORD#9;
                            ELSE wPulse := WORD#16#0100; END_IF;
                        6:
                            IF NOT GVL_RobotBridge.xRobotRunning THEN wReject := WORD#9;
                            ELSE wPulse := WORD#16#0400; END_IF;
                        7:
                            wPulse := WORD#16#0800;
                            xLoadSent := FALSE; GVL_RobotBridge.xLoadOperatorConfirmed := FALSE;
                        8:
                            IF GVL_RobotBridge.xRobotRunning OR GVL_RobotBridge.xRobotPaused THEN wReject := WORD#9;
                            ELSIF GVL_RobotBridge.xRobotAlarm THEN wPulse := WORD#16#0200; END_IF;
                        END_CASE;
                        IF wReject = WORD#0 THEN
                            xHasControlledRobot := TRUE;
                            IF wPulse <> WORD#0 THEN
                                uiStep := UINT#10; xNewAction := TRUE;
                                xRunningSeen := FALSE;
                                wAckResult := WORD#1;
                            END_IF;
                        END_IF;
                    END_IF;
                ELSE
                    CASE WORD_TO_UINT(wCmd) OF
                    9: // Logout only after stop and disable.
                        IF NOT GVL_RobotBridge.xRobotLinkOK OR NOT xTerminalStop
                           OR GVL_RobotBridge.xRobotEnabled THEN wReject := WORD#9;
                        ELSE
                            GVL_RobotBridge.xHostRegistered := FALSE;
                            GVL_RobotBridge.xHostAlive := FALSE;
                            udiOwner := UDINT#0; xHasControlledRobot := FALSE;
                            GVL_RobotBridge.xLoadOperatorConfirmed := FALSE;
                        END_IF;
                    10: // Select coordinates vs AO21..32; no motion request.
                        IF wParam > WORD#1 THEN wReject := WORD#8;
                        ELSIF NOT GVL_RobotBridge.xCommissioned OR NOT GVL_RobotBridge.xRemotePermit
                              OR NOT GVL_RobotBridge.xRobotLinkOK OR NOT xTerminalStop THEN wReject := WORD#9;
                        ELSE xCoordinates := wParam = WORD#1;
                             wAckResult := WORD#3; // Selection sent; no separate selector feedback.
                        END_IF;
                    11: // Explicitly rearm the communications stop latch, never automatic.
                        IF NOT GVL_RobotBridge.xCommissioned OR NOT GVL_RobotBridge.xGdiProgramMappingConfirmed
                           OR NOT GVL_RobotBridge.xRemotePermit
                           OR NOT GVL_RobotBridge.xRobotLinkOK OR NOT xTerminalStop
                           OR GVL_RobotBridge.xRobotEmergency THEN wReject := WORD#9;
                        ELSE
                            GVL_RobotBridge.xStopInterlock := FALSE;
                            xHasControlledRobot := FALSE; xLoadSent := FALSE;
                            GVL_RobotBridge.xLoadOperatorConfirmed := FALSE;
                        END_IF;
                    12: // Operator has CHECKED the actually loaded program on the pendant.
                        IF GVL_FileBridge.xFixedUpdateBusy THEN wReject := WORD#9;
                        ELSIF NOT xLoadSent OR NOT GVL_RobotBridge.xGdiProgramMappingConfirmed
                           OR (wParam <> UINT_TO_WORD(uiSelectedProgram))
                           OR NOT GVL_RobotBridge.xCommissioned OR NOT GVL_RobotBridge.xRemotePermit
                           OR NOT GVL_RobotBridge.xRobotLinkOK OR NOT xTerminalStop
                           OR GVL_RobotBridge.xRobotAlarm OR GVL_RobotBridge.xStopInterlock THEN wReject := WORD#9;
                        ELSE GVL_RobotBridge.xLoadOperatorConfirmed := TRUE;
                        END_IF;
                    ELSE wReject := WORD#8;
                    END_CASE;
                END_IF;
                IF wReject <> WORD#0 THEN
                    wAckResult := WORD#4; wAckError := wReject;
                END_IF;
            END_IF;
        END_IF;
    END_IF;
    IF wReject <> WORD#0 THEN
        udiRejectedSeq := udiRequest; wLastReject := wReject;
    END_IF;
END_IF;

// ----- Pulse timing: each phase owns a separate timer -----
fbLowBefore(IN := (uiStep = UINT#10) AND NOT xNewAction, PT := T#500ms);
fbPulse(IN := (uiStep = UINT#20) AND NOT xNewAction, PT := T#500ms);
fbLowAfter(IN := (uiStep = UINT#30) AND NOT xNewAction, PT := T#500ms);
fbActionTimeout(IN := (uiStep <> UINT#0) AND NOT xNewAction, PT := T#10s);
IF (wAckCmd = WORD#5) AND (uiStep >= UINT#20)
   AND GVL_RobotBridge.xRobotLinkOK AND GVL_RobotBridge.xRobotRunning THEN
    xRunningSeen := TRUE;
END_IF;
CASE uiStep OF
10: IF fbLowBefore.Q THEN uiStep := UINT#20; END_IF;
20: IF fbPulse.Q THEN uiStep := UINT#30; END_IF;
30: IF fbLowAfter.Q THEN uiStep := UINT#40; END_IF;
40:
    xConfirmed := FALSE;
    CASE WORD_TO_UINT(wAckCmd) OF
    2: xConfirmed := GVL_RobotBridge.xRobotEnabled;
    3: xConfirmed := NOT GVL_RobotBridge.xRobotEnabled;
    4: // The supplied standard word has NO dedicated load-complete bit.
        xLoadSent := TRUE; wAckResult := WORD#3; uiStep := UINT#0;
    5: xConfirmed := xRunningSeen;
    6: xConfirmed := GVL_RobotBridge.xRobotPaused AND NOT GVL_RobotBridge.xRobotRunning;
    7: xConfirmed := xTerminalStop;
    8: xConfirmed := NOT GVL_RobotBridge.xRobotAlarm;
    END_CASE;
    IF xConfirmed AND GVL_RobotBridge.xRobotLinkOK THEN
        wAckResult := WORD#2; wAckError := WORD#0; uiStep := UINT#0;
    END_IF;
END_CASE;
IF fbActionTimeout.Q AND (uiStep <> UINT#0) THEN
    uiStep := UINT#0; wAckResult := WORD#5; wAckError := WORD#10;
    GVL_RobotBridge.xStopInterlock := TRUE;
    GVL_RobotBridge.xLoadOperatorConfirmed := FALSE;
END_IF;

// ----- Single writer: FC16 offset 0, TWO consecutive WORDs -----
// aRobotTx[0] owns DI33..48; [1] owns DI49..64. No other writer.
// DI33..36 remain zero: remove legacy one-hot bindings before commissioning.
// DI49 is GDI bit0, DI56 bit7; DI57..64 remain zero.
// Program number settles for 500 ms BEFORE the load rising edge.
GVL_RobotBridge.wRobotTxControl := WORD#0;
IF GVL_RobotBridge.xCommissioned THEN
    IF xCoordinates THEN
        GVL_RobotBridge.wRobotTxControl := GVL_RobotBridge.wRobotTxControl OR WORD#16#1000;
    END_IF;
    IF uiStep = UINT#20 THEN
        GVL_RobotBridge.wRobotTxControl := GVL_RobotBridge.wRobotTxControl OR wPulse;
    END_IF;
    IF GVL_RobotBridge.xStopInterlock THEN
        GVL_RobotBridge.wRobotTxControl := WORD#16#0800;
        IF xCoordinates THEN
            GVL_RobotBridge.wRobotTxControl := GVL_RobotBridge.wRobotTxControl OR WORD#16#1000;
        END_IF;
    END_IF;
END_IF;
GVL_RobotBridge.aRobotTx[0] := GVL_RobotBridge.wRobotTxControl;
GVL_RobotBridge.aRobotTx[1] := WORD#0;
IF GVL_RobotBridge.xCommissioned AND GVL_RobotBridge.xGdiProgramMappingConfirmed THEN
    GVL_RobotBridge.aRobotTx[1] := UINT_TO_WORD(uiSelectedProgram) AND WORD#16#00FF;
END_IF;
GVL_RobotBridge.xBusy := uiStep <> UINT#0;

// ----- PC status: HR300..363, exclusively written here -----
FOR i := 0 TO 63 DO GVL_RobotBridge.aHostStatus[i] := WORD#0; END_FOR;
IF wPlcHb = WORD#16#FFFF THEN wPlcHb := WORD#0;
ELSE wPlcHb := UINT_TO_WORD(WORD_TO_UINT(wPlcHb) + UINT#1); END_IF;
wFlags := WORD#1;
IF GVL_RobotBridge.xRobotLinkOK THEN wFlags := wFlags OR WORD#16#0002; END_IF;
IF GVL_RobotBridge.xRemotePermit THEN wFlags := wFlags OR WORD#16#0004; END_IF;
IF GVL_RobotBridge.xHostRegistered THEN wFlags := wFlags OR WORD#16#0008; END_IF;
IF GVL_RobotBridge.xHostAlive THEN wFlags := wFlags OR WORD#16#0010; END_IF;
IF GVL_RobotBridge.xBusy THEN wFlags := wFlags OR WORD#16#0020; END_IF;
IF GVL_RobotBridge.xCommissioned THEN wFlags := wFlags OR WORD#16#0040; END_IF;
IF xCoordinates THEN wFlags := wFlags OR WORD#16#0080; END_IF;
IF GVL_RobotBridge.xStopInterlock THEN wFlags := wFlags OR WORD#16#0100; END_IF;
IF GVL_RobotBridge.xLoadOperatorConfirmed THEN wFlags := wFlags OR WORD#16#0200; END_IF;
GVL_RobotBridge.aHostStatus[0] := WORD#16#4D42;
GVL_RobotBridge.aHostStatus[1] := WORD#2;
IF GVL_RobotBridge.xGdiProgramMappingConfirmed THEN wFlags := wFlags OR WORD#16#0400; END_IF;
GVL_RobotBridge.aHostStatus[2] := wFlags;
GVL_RobotBridge.aHostStatus[3] := UINT_TO_WORD(uiStep);
GVL_RobotBridge.aHostStatus[4] := UDINT_TO_WORD(SHR(udiAckSeq, 16));
GVL_RobotBridge.aHostStatus[5] := UDINT_TO_WORD(udiAckSeq AND UDINT#65535);
GVL_RobotBridge.aHostStatus[6] := wAckCmd;
GVL_RobotBridge.aHostStatus[7] := wAckResult;
GVL_RobotBridge.aHostStatus[8] := wAckError;
GVL_RobotBridge.aHostStatus[9] := wLastHostHb;
GVL_RobotBridge.aHostStatus[10] := UDINT_TO_WORD(SHR(GVL_RobotBridgeRetain.udiBootCounter, 16));
GVL_RobotBridge.aHostStatus[11] := UDINT_TO_WORD(GVL_RobotBridgeRetain.udiBootCounter AND UDINT#65535);
GVL_RobotBridge.aHostStatus[12] := wPlcHb;
GVL_RobotBridge.aHostStatus[13] := UINT_TO_WORD(uiSelectedProgram);
GVL_RobotBridge.aHostStatus[14] := GVL_RobotBridge.wRobotTxControl;
GVL_RobotBridge.aHostStatus[15] := UDINT_TO_WORD(SHR(udiOwner, 16));
GVL_RobotBridge.aHostStatus[16] := UDINT_TO_WORD(udiOwner AND UDINT#65535);
GVL_RobotBridge.aHostStatus[17] := GVL_RobotBridge.aRobotRx[0];
IF NOT GVL_RobotBridge.xRobotLinkOK THEN GVL_RobotBridge.aHostStatus[18] := WORD#0;
ELSIF GVL_RobotBridge.xRobotEmergency THEN GVL_RobotBridge.aHostStatus[18] := WORD#5;
ELSIF GVL_RobotBridge.xRobotAlarm THEN GVL_RobotBridge.aHostStatus[18] := WORD#4;
ELSIF GVL_RobotBridge.xRobotPaused THEN GVL_RobotBridge.aHostStatus[18] := WORD#3;
ELSIF GVL_RobotBridge.xRobotRunning THEN GVL_RobotBridge.aHostStatus[18] := WORD#2;
ELSIF xTerminalStop THEN GVL_RobotBridge.aHostStatus[18] := WORD#1;
END_IF;
FOR i := 0 TO 31 DO
    GVL_RobotBridge.aHostStatus[20 + i] := GVL_RobotBridge.aRobotRx[i];
END_FOR;
GVL_RobotBridge.aHostStatus[52] := UDINT_TO_WORD(SHR(udiRejectedSeq, 16));
GVL_RobotBridge.aHostStatus[53] := UDINT_TO_WORD(udiRejectedSeq AND UDINT#65535);
GVL_RobotBridge.aHostStatus[54] := wLastReject;
GVL_RobotBridge.aHostStatus[55] := UDINT_TO_WORD(SHR(udiInterruptedSeq, 16));
GVL_RobotBridge.aHostStatus[56] := UDINT_TO_WORD(udiInterruptedSeq AND UDINT#65535);
GVL_RobotBridge.aHostStatus[62] := wHbCount;

// V2 capability block; desired program word is NOT robot readback.
GVL_RobotBridge.aHostStatus[57] := WORD#1; // selection mode: 1 = GDI8
GVL_RobotBridge.aHostStatus[58] := WORD#255; // maximum program number
GVL_RobotBridge.aHostStatus[59] := GVL_RobotBridge.aRobotTx[1];
GVL_RobotBridge.aHostStatus[60] := WORD#49; // first GDI DI (bit0)
GVL_RobotBridge.aHostStatus[61] := WORD#56; // last GDI DI (bit7)
GVL_RobotBridge.aHostStatus[63] := WORD#2; // robot FC16 write word count
END_PROGRAM
